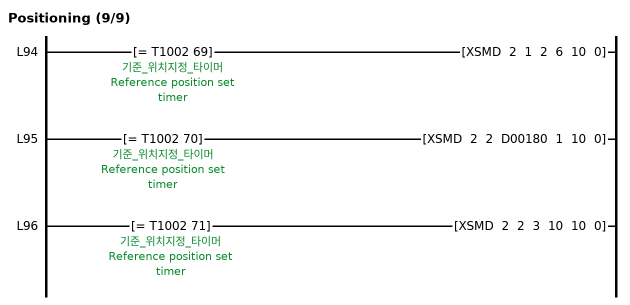
[picture p24: Positioning rungs L94-L96]
; L94
LOAD=     T1002 69	// 기준_위치지정_타이머 Reference position set timer
XSMD      2 1 2 6 10 0
; L95
LOAD=     T1002 70	// 기준_위치지정_타이머 Reference position set timer
XSMD      2 2 D00180 1 10 0
; L96
LOAD=     T1002 71	// 기준_위치지정_타이머 Reference position set timer
XSMD      2 2 3 10 10 0

PROGRAM PosItion_Switch (task: 스캔 프로그램)

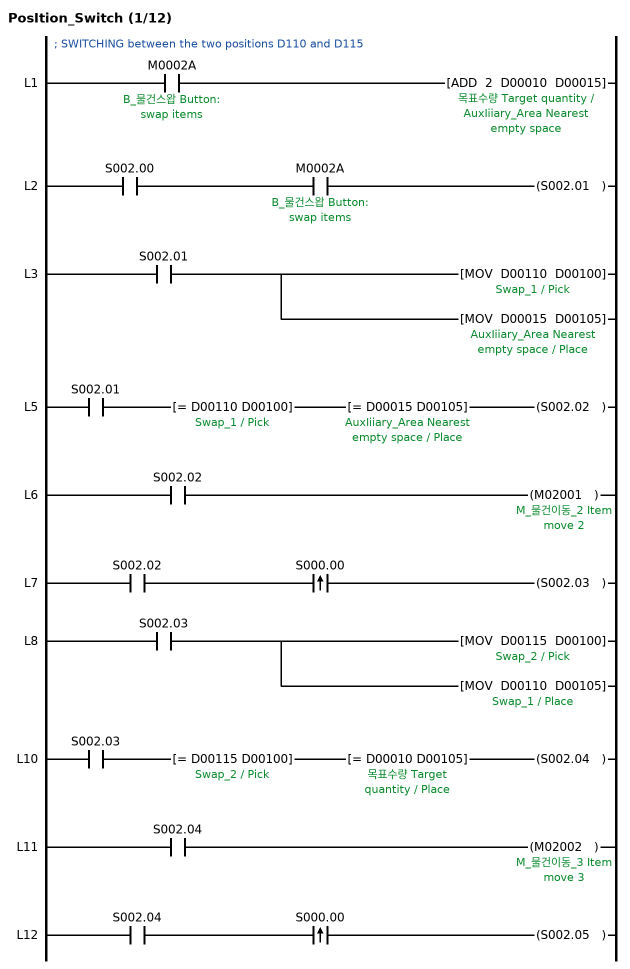
// SWITCHING between the two positions D110 and D115
; L1
LOAD      M0002A	// B_물건스왑 Button: swap items
ADD       2 D00010 D00015	// 목표수량 Target quantity / AuxIiiary_Area Nearest empty space
; L2
LOAD      S002.00
AND       M0002A	// B_물건스왑 Button: swap items
OUT       S002.01
; L3
LOAD      S002.01
MOV       D00110 D00100	// Swap_1 / Pick
MOV       D00015 D00105	// AuxIiiary_Area Nearest empty space / Place
; L5
LOAD      S002.01
AND=      D00110 D00100	// Swap_1 / Pick
AND=      D00015 D00105	// AuxIiiary_Area Nearest empty space / Place
OUT       S002.02
; L6
LOAD      S002.02
OUT       M02001	// M_물건이동_2 Item move 2
; L7
LOAD      S002.02
ANDP      S000.00
OUT       S002.03
; L8
LOAD      S002.03
MOV       D00115 D00100	// Swap_2 / Pick
MOV       D00110 D00105	// Swap_1 / Place
; L10
LOAD      S002.03
AND=      D00115 D00100	// Swap_2 / Pick
AND=      D00010 D00105	// 목표수량 Target quantity / Place
OUT       S002.04
; L11
LOAD      S002.04
OUT       M02002	// M_물건이동_3 Item move 3
; L12
LOAD      S002.04
ANDP      S000.00
OUT       S002.05

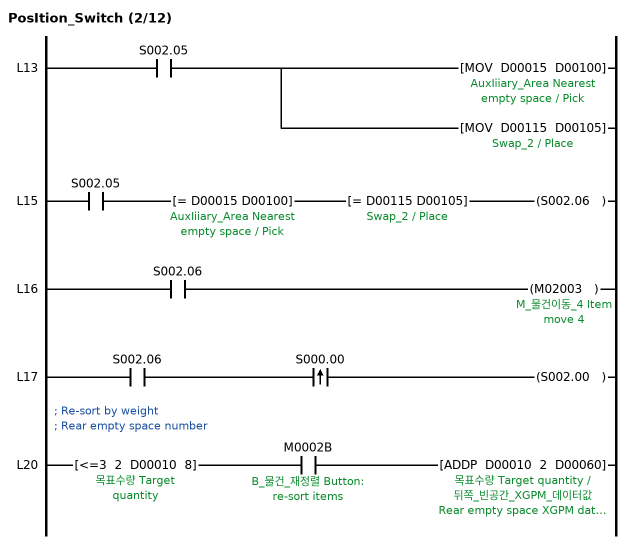
; L13
LOAD      S002.05
MOV       D00015 D00100	// AuxIiiary_Area Nearest empty space / Pick
MOV       D00115 D00105	// Swap_2 / Place
; L15
LOAD      S002.05
AND=      D00015 D00100	// AuxIiiary_Area Nearest empty space / Pick
AND=      D00115 D00105	// Swap_2 / Place
OUT       S002.06
; L16
LOAD      S002.06
OUT       M02003	// M_물건이동_4 Item move 4
; L17
LOAD      S002.06
ANDP      S000.00
OUT       S002.00
// Re-sort by weight
// Rear empty space number
; L20
LOAD<=3   2 D00010 8	// 목표수량 Target quantity
AND       M0002B	// B_물건_재정렬 Button: re-sort items
ADDP      D00010 2 D00060	// 목표수량 Target quantity / 뒤쪽_빈공간_XGPM_데이터값 Rear empty space XGPM data value

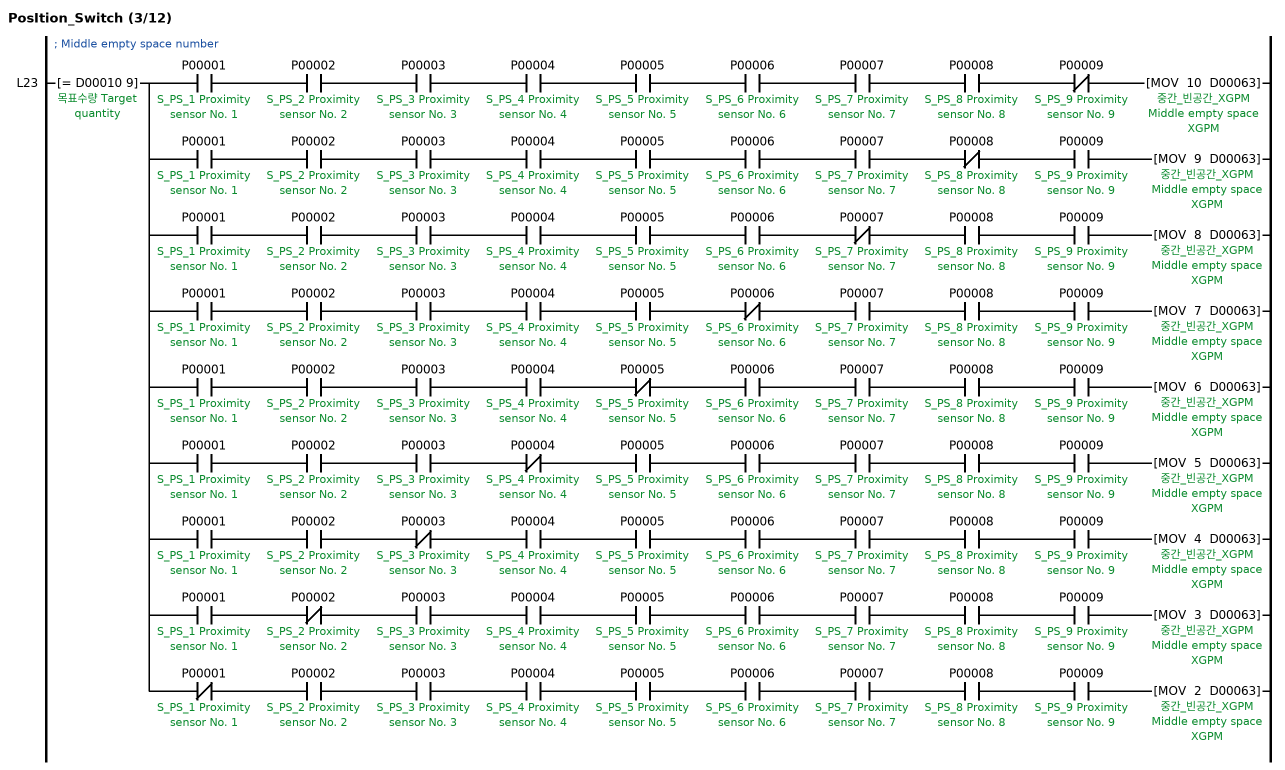
// Middle empty space number
; L23
LOAD=     D00010 9	// 목표수량 Target quantity
MPUSH
AND       P00001	// S_PS_1 Proximity sensor No. 1
AND       P00002	// S_PS_2 Proximity sensor No. 2
AND       P00003	// S_PS_3 Proximity sensor No. 3
AND       P00004	// S_PS_4 Proximity sensor No. 4
AND       P00005	// S_PS_5 Proximity sensor No. 5
AND       P00006	// S_PS_6 Proximity sensor No. 6
AND       P00007	// S_PS_7 Proximity sensor No. 7
AND       P00008	// S_PS_8 Proximity sensor No. 8
AND NOT   P00009	// S_PS_9 Proximity sensor No. 9
MOV       10 D00063	// 중간_빈공간_XGPM Middle empty space XGPM
MLOAD
AND       P00001	// S_PS_1 Proximity sensor No. 1
AND       P00002	// S_PS_2 Proximity sensor No. 2
AND       P00003	// S_PS_3 Proximity sensor No. 3
AND       P00004	// S_PS_4 Proximity sensor No. 4
AND       P00005	// S_PS_5 Proximity sensor No. 5
AND       P00006	// S_PS_6 Proximity sensor No. 6
AND       P00007	// S_PS_7 Proximity sensor No. 7
AND NOT   P00008	// S_PS_8 Proximity sensor No. 8
AND       P00009	// S_PS_9 Proximity sensor No. 9
MOV       9 D00063	// 중간_빈공간_XGPM Middle empty space XGPM
MLOAD
AND       P00001	// S_PS_1 Proximity sensor No. 1
AND       P00002	// S_PS_2 Proximity sensor No. 2
AND       P00003	// S_PS_3 Proximity sensor No. 3
AND       P00004	// S_PS_4 Proximity sensor No. 4
AND       P00005	// S_PS_5 Proximity sensor No. 5
AND       P00006	// S_PS_6 Proximity sensor No. 6
AND NOT   P00007	// S_PS_7 Proximity sensor No. 7
AND       P00008	// S_PS_8 Proximity sensor No. 8
AND       P00009	// S_PS_9 Proximity sensor No. 9
MOV       8 D00063	// 중간_빈공간_XGPM Middle empty space XGPM
MLOAD
AND       P00001	// S_PS_1 Proximity sensor No. 1
AND       P00002	// S_PS_2 Proximity sensor No. 2
AND       P00003	// S_PS_3 Proximity sensor No. 3
AND       P00004	// S_PS_4 Proximity sensor No. 4
AND       P00005	// S_PS_5 Proximity sensor No. 5
AND NOT   P00006	// S_PS_6 Proximity sensor No. 6
AND       P00007	// S_PS_7 Proximity sensor No. 7
AND       P00008	// S_PS_8 Proximity sensor No. 8
AND       P00009	// S_PS_9 Proximity sensor No. 9
MOV       7 D00063	// 중간_빈공간_XGPM Middle empty space XGPM
MLOAD
AND       P00001	// S_PS_1 Proximity sensor No. 1
AND       P00002	// S_PS_2 Proximity sensor No. 2
AND       P00003	// S_PS_3 Proximity sensor No. 3
AND       P00004	// S_PS_4 Proximity sensor No. 4
AND NOT   P00005	// S_PS_5 Proximity sensor No. 5
AND       P00006	// S_PS_6 Proximity sensor No. 6
AND       P00007	// S_PS_7 Proximity sensor No. 7
AND       P00008	// S_PS_8 Proximity sensor No. 8
AND       P00009	// S_PS_9 Proximity sensor No. 9
MOV       6 D00063	// 중간_빈공간_XGPM Middle empty space XGPM
MLOAD
AND       P00001	// S_PS_1 Proximity sensor No. 1
AND       P00002	// S_PS_2 Proximity sensor No. 2
AND       P00003	// S_PS_3 Proximity sensor No. 3
AND NOT   P00004	// S_PS_4 Proximity sensor No. 4
AND       P00005	// S_PS_5 Proximity sensor No. 5
AND       P00006	// S_PS_6 Proximity sensor No. 6
AND       P00007	// S_PS_7 Proximity sensor No. 7
AND       P00008	// S_PS_8 Proximity sensor No. 8
AND       P00009	// S_PS_9 Proximity sensor No. 9
MOV       5 D00063	// 중간_빈공간_XGPM Middle empty space XGPM
MLOAD
AND       P00001	// S_PS_1 Proximity sensor No. 1
AND       P00002	// S_PS_2 Proximity sensor No. 2
AND NOT   P00003	// S_PS_3 Proximity sensor No. 3
AND       P00004	// S_PS_4 Proximity sensor No. 4
AND       P00005	// S_PS_5 Proximity sensor No. 5
AND       P00006	// S_PS_6 Proximity sensor No. 6
AND       P00007	// S_PS_7 Proximity sensor No. 7
AND       P00008	// S_PS_8 Proximity sensor No. 8
AND       P00009	// S_PS_9 Proximity sensor No. 9
MOV       4 D00063	// 중간_빈공간_XGPM Middle empty space XGPM
MLOAD
AND       P00001	// S_PS_1 Proximity sensor No. 1
AND NOT   P00002	// S_PS_2 Proximity sensor No. 2
AND       P00003	// S_PS_3 Proximity sensor No. 3
AND       P00004	// S_PS_4 Proximity sensor No. 4
AND       P00005	// S_PS_5 Proximity sensor No. 5
AND       P00006	// S_PS_6 Proximity sensor No. 6
AND       P00007	// S_PS_7 Proximity sensor No. 7
AND       P00008	// S_PS_8 Proximity sensor No. 8
AND       P00009	// S_PS_9 Proximity sensor No. 9
MOV       3 D00063	// 중간_빈공간_XGPM Middle empty space XGPM
MPOP
AND NOT   P00001	// S_PS_1 Proximity sensor No. 1
AND       P00002	// S_PS_2 Proximity sensor No. 2
AND       P00003	// S_PS_3 Proximity sensor No. 3
AND       P00004	// S_PS_4 Proximity sensor No. 4
AND       P00005	// S_PS_5 Proximity sensor No. 5
AND       P00006	// S_PS_6 Proximity sensor No. 6
AND       P00007	// S_PS_7 Proximity sensor No. 7
AND       P00008	// S_PS_8 Proximity sensor No. 8
AND       P00009	// S_PS_9 Proximity sensor No. 9
MOV       2 D00063	// 중간_빈공간_XGPM Middle empty space XGPM

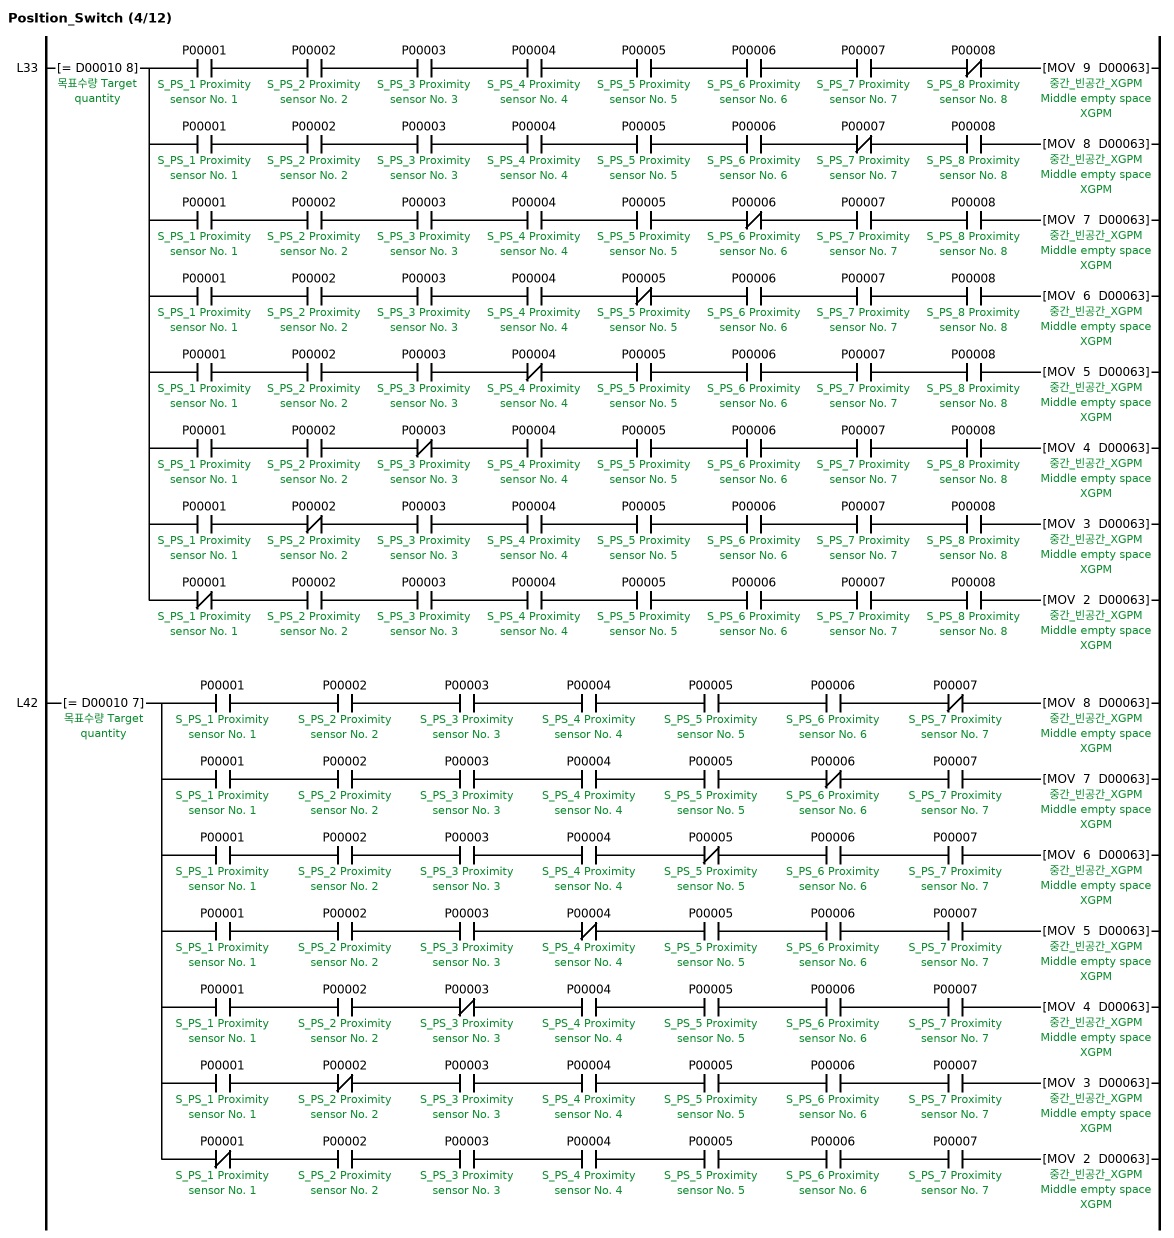
; L33
LOAD=     D00010 8	// 목표수량 Target quantity
MPUSH
AND       P00001	// S_PS_1 Proximity sensor No. 1
AND       P00002	// S_PS_2 Proximity sensor No. 2
AND       P00003	// S_PS_3 Proximity sensor No. 3
AND       P00004	// S_PS_4 Proximity sensor No. 4
AND       P00005	// S_PS_5 Proximity sensor No. 5
AND       P00006	// S_PS_6 Proximity sensor No. 6
AND       P00007	// S_PS_7 Proximity sensor No. 7
AND NOT   P00008	// S_PS_8 Proximity sensor No. 8
MOV       9 D00063	// 중간_빈공간_XGPM Middle empty space XGPM
MLOAD
AND       P00001	// S_PS_1 Proximity sensor No. 1
AND       P00002	// S_PS_2 Proximity sensor No. 2
AND       P00003	// S_PS_3 Proximity sensor No. 3
AND       P00004	// S_PS_4 Proximity sensor No. 4
AND       P00005	// S_PS_5 Proximity sensor No. 5
AND       P00006	// S_PS_6 Proximity sensor No. 6
AND NOT   P00007	// S_PS_7 Proximity sensor No. 7
AND       P00008	// S_PS_8 Proximity sensor No. 8
MOV       8 D00063	// 중간_빈공간_XGPM Middle empty space XGPM
MLOAD
AND       P00001	// S_PS_1 Proximity sensor No. 1
AND       P00002	// S_PS_2 Proximity sensor No. 2
AND       P00003	// S_PS_3 Proximity sensor No. 3
AND       P00004	// S_PS_4 Proximity sensor No. 4
AND       P00005	// S_PS_5 Proximity sensor No. 5
AND NOT   P00006	// S_PS_6 Proximity sensor No. 6
AND       P00007	// S_PS_7 Proximity sensor No. 7
AND       P00008	// S_PS_8 Proximity sensor No. 8
MOV       7 D00063	// 중간_빈공간_XGPM Middle empty space XGPM
MLOAD
AND       P00001	// S_PS_1 Proximity sensor No. 1
AND       P00002	// S_PS_2 Proximity sensor No. 2
AND       P00003	// S_PS_3 Proximity sensor No. 3
AND       P00004	// S_PS_4 Proximity sensor No. 4
AND NOT   P00005	// S_PS_5 Proximity sensor No. 5
AND       P00006	// S_PS_6 Proximity sensor No. 6
AND       P00007	// S_PS_7 Proximity sensor No. 7
AND       P00008	// S_PS_8 Proximity sensor No. 8
MOV       6 D00063	// 중간_빈공간_XGPM Middle empty space XGPM
MLOAD
AND       P00001	// S_PS_1 Proximity sensor No. 1
AND       P00002	// S_PS_2 Proximity sensor No. 2
AND       P00003	// S_PS_3 Proximity sensor No. 3
AND NOT   P00004	// S_PS_4 Proximity sensor No. 4
AND       P00005	// S_PS_5 Proximity sensor No. 5
AND       P00006	// S_PS_6 Proximity sensor No. 6
AND       P00007	// S_PS_7 Proximity sensor No. 7
AND       P00008	// S_PS_8 Proximity sensor No. 8
MOV       5 D00063	// 중간_빈공간_XGPM Middle empty space XGPM
MLOAD
AND       P00001	// S_PS_1 Proximity sensor No. 1
AND       P00002	// S_PS_2 Proximity sensor No. 2
AND NOT   P00003	// S_PS_3 Proximity sensor No. 3
AND       P00004	// S_PS_4 Proximity sensor No. 4
AND       P00005	// S_PS_5 Proximity sensor No. 5
AND       P00006	// S_PS_6 Proximity sensor No. 6
AND       P00007	// S_PS_7 Proximity sensor No. 7
AND       P00008	// S_PS_8 Proximity sensor No. 8
MOV       4 D00063	// 중간_빈공간_XGPM Middle empty space XGPM
MLOAD
AND       P00001	// S_PS_1 Proximity sensor No. 1
AND NOT   P00002	// S_PS_2 Proximity sensor No. 2
AND       P00003	// S_PS_3 Proximity sensor No. 3
AND       P00004	// S_PS_4 Proximity sensor No. 4
AND       P00005	// S_PS_5 Proximity sensor No. 5
AND       P00006	// S_PS_6 Proximity sensor No. 6
AND       P00007	// S_PS_7 Proximity sensor No. 7
AND       P00008	// S_PS_8 Proximity sensor No. 8
MOV       3 D00063	// 중간_빈공간_XGPM Middle empty space XGPM
MPOP
AND NOT   P00001	// S_PS_1 Proximity sensor No. 1
AND       P00002	// S_PS_2 Proximity sensor No. 2
AND       P00003	// S_PS_3 Proximity sensor No. 3
AND       P00004	// S_PS_4 Proximity sensor No. 4
AND       P00005	// S_PS_5 Proximity sensor No. 5
AND       P00006	// S_PS_6 Proximity sensor No. 6
AND       P00007	// S_PS_7 Proximity sensor No. 7
AND       P00008	// S_PS_8 Proximity sensor No. 8
MOV       2 D00063	// 중간_빈공간_XGPM Middle empty space XGPM
; L42
LOAD=     D00010 7	// 목표수량 Target quantity
MPUSH
AND       P00001	// S_PS_1 Proximity sensor No. 1
AND       P00002	// S_PS_2 Proximity sensor No. 2
AND       P00003	// S_PS_3 Proximity sensor No. 3
AND       P00004	// S_PS_4 Proximity sensor No. 4
AND       P00005	// S_PS_5 Proximity sensor No. 5
AND       P00006	// S_PS_6 Proximity sensor No. 6
AND NOT   P00007	// S_PS_7 Proximity sensor No. 7
MOV       8 D00063	// 중간_빈공간_XGPM Middle empty space XGPM
MLOAD
AND       P00001	// S_PS_1 Proximity sensor No. 1
AND       P00002	// S_PS_2 Proximity sensor No. 2
AND       P00003	// S_PS_3 Proximity sensor No. 3
AND       P00004	// S_PS_4 Proximity sensor No. 4
AND       P00005	// S_PS_5 Proximity sensor No. 5
AND NOT   P00006	// S_PS_6 Proximity sensor No. 6
AND       P00007	// S_PS_7 Proximity sensor No. 7
MOV       7 D00063	// 중간_빈공간_XGPM Middle empty space XGPM
MLOAD
AND       P00001	// S_PS_1 Proximity sensor No. 1
AND       P00002	// S_PS_2 Proximity sensor No. 2
AND       P00003	// S_PS_3 Proximity sensor No. 3
AND       P00004	// S_PS_4 Proximity sensor No. 4
AND NOT   P00005	// S_PS_5 Proximity sensor No. 5
AND       P00006	// S_PS_6 Proximity sensor No. 6
AND       P00007	// S_PS_7 Proximity sensor No. 7
MOV       6 D00063	// 중간_빈공간_XGPM Middle empty space XGPM
MLOAD
AND       P00001	// S_PS_1 Proximity sensor No. 1
AND       P00002	// S_PS_2 Proximity sensor No. 2
AND       P00003	// S_PS_3 Proximity sensor No. 3
AND NOT   P00004	// S_PS_4 Proximity sensor No. 4
AND       P00005	// S_PS_5 Proximity sensor No. 5
AND       P00006	// S_PS_6 Proximity sensor No. 6
AND       P00007	// S_PS_7 Proximity sensor No. 7
MOV       5 D00063	// 중간_빈공간_XGPM Middle empty space XGPM
MLOAD
AND       P00001	// S_PS_1 Proximity sensor No. 1
AND       P00002	// S_PS_2 Proximity sensor No. 2
AND NOT   P00003	// S_PS_3 Proximity sensor No. 3
AND       P00004	// S_PS_4 Proximity sensor No. 4
AND       P00005	// S_PS_5 Proximity sensor No. 5
AND       P00006	// S_PS_6 Proximity sensor No. 6
AND       P00007	// S_PS_7 Proximity sensor No. 7
MOV       4 D00063	// 중간_빈공간_XGPM Middle empty space XGPM
MLOAD
AND       P00001	// S_PS_1 Proximity sensor No. 1
AND NOT   P00002	// S_PS_2 Proximity sensor No. 2
AND       P00003	// S_PS_3 Proximity sensor No. 3
AND       P00004	// S_PS_4 Proximity sensor No. 4
AND       P00005	// S_PS_5 Proximity sensor No. 5
AND       P00006	// S_PS_6 Proximity sensor No. 6
AND       P00007	// S_PS_7 Proximity sensor No. 7
MOV       3 D00063	// 중간_빈공간_XGPM Middle empty space XGPM
MPOP
AND NOT   P00001	// S_PS_1 Proximity sensor No. 1
AND       P00002	// S_PS_2 Proximity sensor No. 2
AND       P00003	// S_PS_3 Proximity sensor No. 3
AND       P00004	// S_PS_4 Proximity sensor No. 4
AND       P00005	// S_PS_5 Proximity sensor No. 5
AND       P00006	// S_PS_6 Proximity sensor No. 6
AND       P00007	// S_PS_7 Proximity sensor No. 7
MOV       2 D00063	// 중간_빈공간_XGPM Middle empty space XGPM

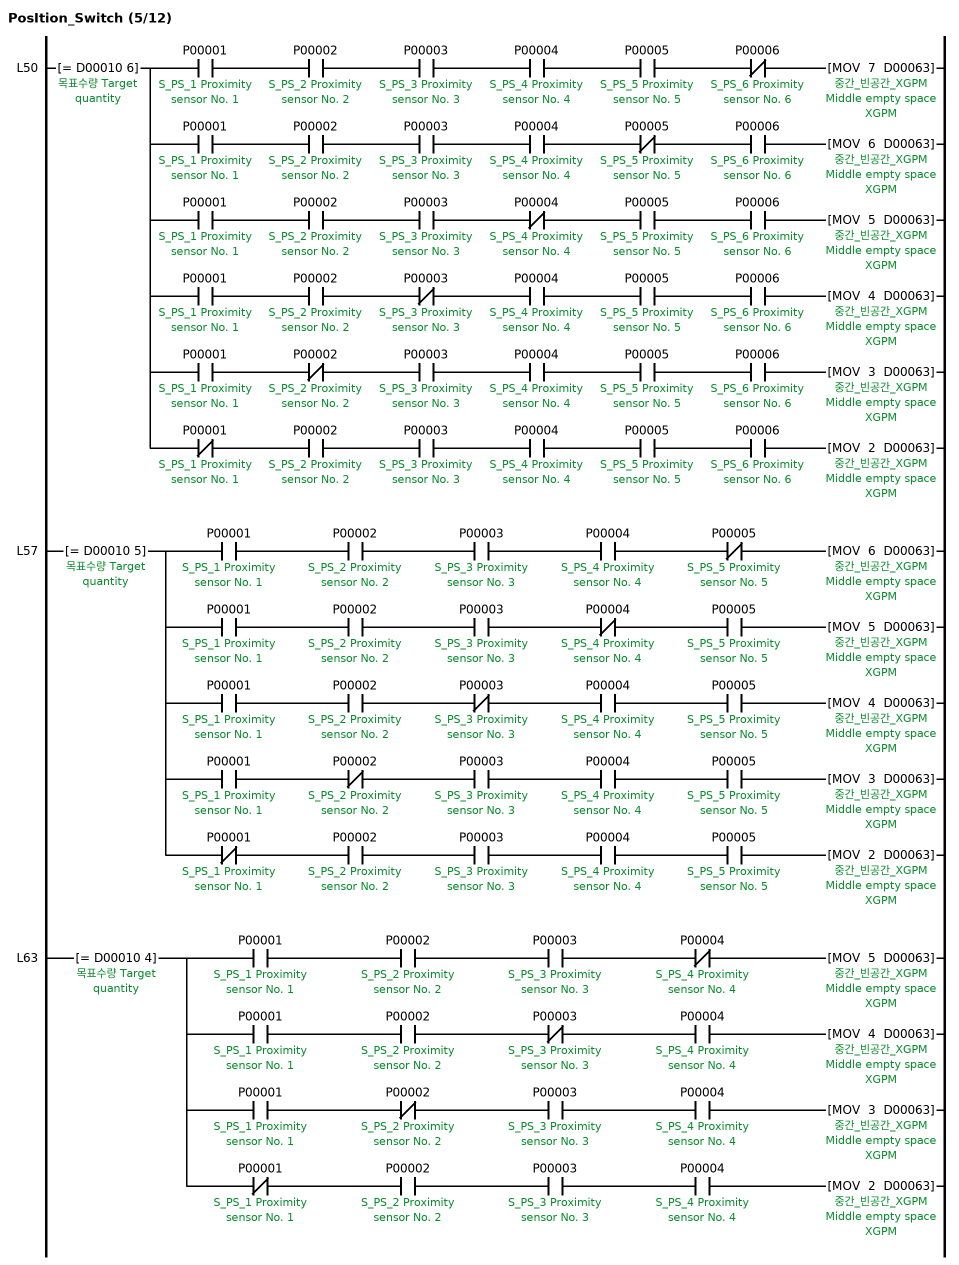
; L50
LOAD=     D00010 6	// 목표수량 Target quantity
MPUSH
AND       P00001	// S_PS_1 Proximity sensor No. 1
AND       P00002	// S_PS_2 Proximity sensor No. 2
AND       P00003	// S_PS_3 Proximity sensor No. 3
AND       P00004	// S_PS_4 Proximity sensor No. 4
AND       P00005	// S_PS_5 Proximity sensor No. 5
AND NOT   P00006	// S_PS_6 Proximity sensor No. 6
MOV       7 D00063	// 중간_빈공간_XGPM Middle empty space XGPM
MLOAD
AND       P00001	// S_PS_1 Proximity sensor No. 1
AND       P00002	// S_PS_2 Proximity sensor No. 2
AND       P00003	// S_PS_3 Proximity sensor No. 3
AND       P00004	// S_PS_4 Proximity sensor No. 4
AND NOT   P00005	// S_PS_5 Proximity sensor No. 5
AND       P00006	// S_PS_6 Proximity sensor No. 6
MOV       6 D00063	// 중간_빈공간_XGPM Middle empty space XGPM
MLOAD
AND       P00001	// S_PS_1 Proximity sensor No. 1
AND       P00002	// S_PS_2 Proximity sensor No. 2
AND       P00003	// S_PS_3 Proximity sensor No. 3
AND NOT   P00004	// S_PS_4 Proximity sensor No. 4
AND       P00005	// S_PS_5 Proximity sensor No. 5
AND       P00006	// S_PS_6 Proximity sensor No. 6
MOV       5 D00063	// 중간_빈공간_XGPM Middle empty space XGPM
MLOAD
AND       P00001	// S_PS_1 Proximity sensor No. 1
AND       P00002	// S_PS_2 Proximity sensor No. 2
AND NOT   P00003	// S_PS_3 Proximity sensor No. 3
AND       P00004	// S_PS_4 Proximity sensor No. 4
AND       P00005	// S_PS_5 Proximity sensor No. 5
AND       P00006	// S_PS_6 Proximity sensor No. 6
MOV       4 D00063	// 중간_빈공간_XGPM Middle empty space XGPM
MLOAD
AND       P00001	// S_PS_1 Proximity sensor No. 1
AND NOT   P00002	// S_PS_2 Proximity sensor No. 2
AND       P00003	// S_PS_3 Proximity sensor No. 3
AND       P00004	// S_PS_4 Proximity sensor No. 4
AND       P00005	// S_PS_5 Proximity sensor No. 5
AND       P00006	// S_PS_6 Proximity sensor No. 6
MOV       3 D00063	// 중간_빈공간_XGPM Middle empty space XGPM
MPOP
AND NOT   P00001	// S_PS_1 Proximity sensor No. 1
AND       P00002	// S_PS_2 Proximity sensor No. 2
AND       P00003	// S_PS_3 Proximity sensor No. 3
AND       P00004	// S_PS_4 Proximity sensor No. 4
AND       P00005	// S_PS_5 Proximity sensor No. 5
AND       P00006	// S_PS_6 Proximity sensor No. 6
MOV       2 D00063	// 중간_빈공간_XGPM Middle empty space XGPM
; L57
LOAD=     D00010 5	// 목표수량 Target quantity
MPUSH
AND       P00001	// S_PS_1 Proximity sensor No. 1
AND       P00002	// S_PS_2 Proximity sensor No. 2
AND       P00003	// S_PS_3 Proximity sensor No. 3
AND       P00004	// S_PS_4 Proximity sensor No. 4
AND NOT   P00005	// S_PS_5 Proximity sensor No. 5
MOV       6 D00063	// 중간_빈공간_XGPM Middle empty space XGPM
MLOAD
AND       P00001	// S_PS_1 Proximity sensor No. 1
AND       P00002	// S_PS_2 Proximity sensor No. 2
AND       P00003	// S_PS_3 Proximity sensor No. 3
AND NOT   P00004	// S_PS_4 Proximity sensor No. 4
AND       P00005	// S_PS_5 Proximity sensor No. 5
MOV       5 D00063	// 중간_빈공간_XGPM Middle empty space XGPM
MLOAD
AND       P00001	// S_PS_1 Proximity sensor No. 1
AND       P00002	// S_PS_2 Proximity sensor No. 2
AND NOT   P00003	// S_PS_3 Proximity sensor No. 3
AND       P00004	// S_PS_4 Proximity sensor No. 4
AND       P00005	// S_PS_5 Proximity sensor No. 5
MOV       4 D00063	// 중간_빈공간_XGPM Middle empty space XGPM
MLOAD
AND       P00001	// S_PS_1 Proximity sensor No. 1
AND NOT   P00002	// S_PS_2 Proximity sensor No. 2
AND       P00003	// S_PS_3 Proximity sensor No. 3
AND       P00004	// S_PS_4 Proximity sensor No. 4
AND       P00005	// S_PS_5 Proximity sensor No. 5
MOV       3 D00063	// 중간_빈공간_XGPM Middle empty space XGPM
MPOP
AND NOT   P00001	// S_PS_1 Proximity sensor No. 1
AND       P00002	// S_PS_2 Proximity sensor No. 2
AND       P00003	// S_PS_3 Proximity sensor No. 3
AND       P00004	// S_PS_4 Proximity sensor No. 4
AND       P00005	// S_PS_5 Proximity sensor No. 5
MOV       2 D00063	// 중간_빈공간_XGPM Middle empty space XGPM
; L63
LOAD=     D00010 4	// 목표수량 Target quantity
MPUSH
AND       P00001	// S_PS_1 Proximity sensor No. 1
AND       P00002	// S_PS_2 Proximity sensor No. 2
AND       P00003	// S_PS_3 Proximity sensor No. 3
AND NOT   P00004	// S_PS_4 Proximity sensor No. 4
MOV       5 D00063	// 중간_빈공간_XGPM Middle empty space XGPM
MLOAD
AND       P00001	// S_PS_1 Proximity sensor No. 1
AND       P00002	// S_PS_2 Proximity sensor No. 2
AND NOT   P00003	// S_PS_3 Proximity sensor No. 3
AND       P00004	// S_PS_4 Proximity sensor No. 4
MOV       4 D00063	// 중간_빈공간_XGPM Middle empty space XGPM
MLOAD
AND       P00001	// S_PS_1 Proximity sensor No. 1
AND NOT   P00002	// S_PS_2 Proximity sensor No. 2
AND       P00003	// S_PS_3 Proximity sensor No. 3
AND       P00004	// S_PS_4 Proximity sensor No. 4
MOV       3 D00063	// 중간_빈공간_XGPM Middle empty space XGPM
MPOP
AND NOT   P00001	// S_PS_1 Proximity sensor No. 1
AND       P00002	// S_PS_2 Proximity sensor No. 2
AND       P00003	// S_PS_3 Proximity sensor No. 3
AND       P00004	// S_PS_4 Proximity sensor No. 4
MOV       2 D00063	// 중간_빈공간_XGPM Middle empty space XGPM

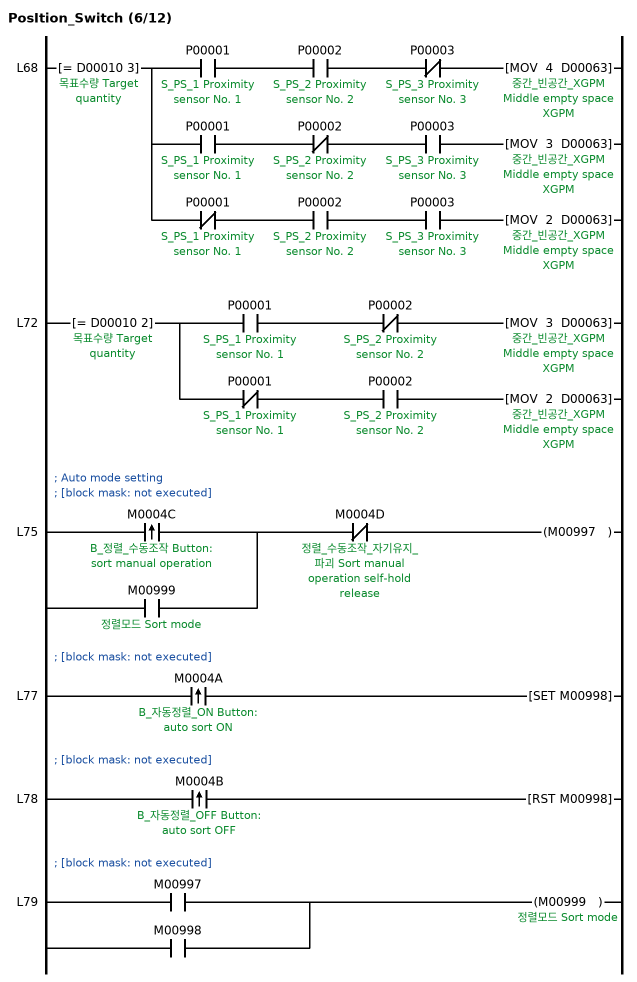
; L68
LOAD=     D00010 3	// 목표수량 Target quantity
MPUSH
AND       P00001	// S_PS_1 Proximity sensor No. 1
AND       P00002	// S_PS_2 Proximity sensor No. 2
AND NOT   P00003	// S_PS_3 Proximity sensor No. 3
MOV       4 D00063	// 중간_빈공간_XGPM Middle empty space XGPM
MLOAD
AND       P00001	// S_PS_1 Proximity sensor No. 1
AND NOT   P00002	// S_PS_2 Proximity sensor No. 2
AND       P00003	// S_PS_3 Proximity sensor No. 3
MOV       3 D00063	// 중간_빈공간_XGPM Middle empty space XGPM
MPOP
AND NOT   P00001	// S_PS_1 Proximity sensor No. 1
AND       P00002	// S_PS_2 Proximity sensor No. 2
AND       P00003	// S_PS_3 Proximity sensor No. 3
MOV       2 D00063	// 중간_빈공간_XGPM Middle empty space XGPM
; L72
LOAD=     D00010 2	// 목표수량 Target quantity
MPUSH
AND       P00001	// S_PS_1 Proximity sensor No. 1
AND NOT   P00002	// S_PS_2 Proximity sensor No. 2
MOV       3 D00063	// 중간_빈공간_XGPM Middle empty space XGPM
MPOP
AND NOT   P00001	// S_PS_1 Proximity sensor No. 1
AND       P00002	// S_PS_2 Proximity sensor No. 2
MOV       2 D00063	// 중간_빈공간_XGPM Middle empty space XGPM
// Auto mode setting
; L75 (block mask: not executed)
LOADP     M0004C	// B_정렬_수동조작 Button: sort manual operation
OR        M00999	// 정렬모드 Sort mode
AND NOT   M0004D	// 정렬_수동조작_자기유지_파괴 Sort manual operation self-hold release
OUT       M00997
; L77 (block mask: not executed)
LOADP     M0004A	// B_자동정렬_ON Button: auto sort ON
SET       M00998
; L78 (block mask: not executed)
LOADP     M0004B	// B_자동정렬_OFF Button: auto sort OFF
RST       M00998
; L79 (block mask: not executed)
LOAD      M00997
OR        M00998
OUT       M00999	// 정렬모드 Sort mode

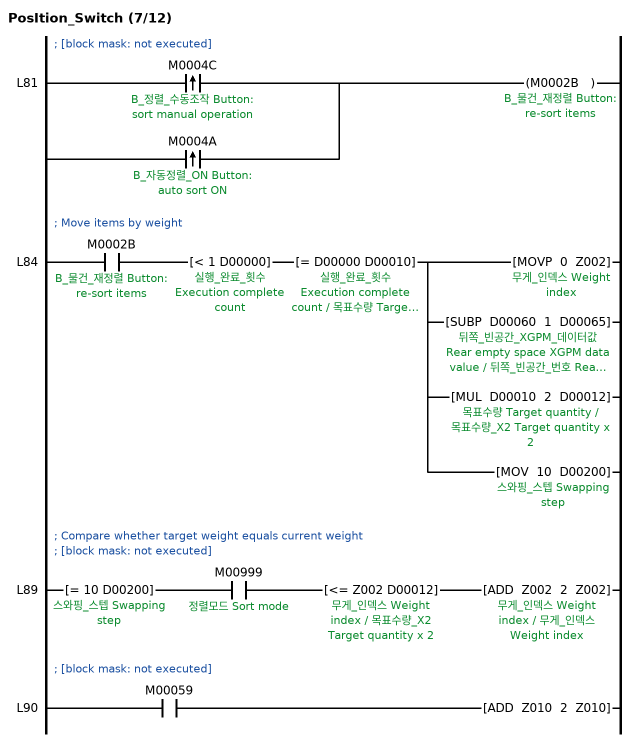
; L81 (block mask: not executed)
LOADP     M0004C	// B_정렬_수동조작 Button: sort manual operation
ORP       M0004A	// B_자동정렬_ON Button: auto sort ON
OUT       M0002B	// B_물건_재정렬 Button: re-sort items
// Move items by weight
; L84
LOAD      M0002B	// B_물건_재정렬 Button: re-sort items
AND<      1 D00000	// 실행_완료_횟수 Execution complete count
AND=      D00000 D00010	// 실행_완료_횟수 Execution complete count / 목표수량 Target quantity
MOVP      0 Z002	// 무게_인덱스 Weight index
SUBP      D00060 1 D00065	// 뒤쪽_빈공간_XGPM_데이터값 Rear empty space XGPM data value / 뒤쪽_빈공간_번호 Rear empty space number
MUL       D00010 2 D00012	// 목표수량 Target quantity / 목표수량_X2 Target quantity x 2
MOV       10 D00200	// 스와핑_스텝 Swapping step
// Compare whether target weight equals current weight
; L89 (block mask: not executed)
LOAD=     10 D00200	// 스와핑_스텝 Swapping step
AND       M00999	// 정렬모드 Sort mode
AND<=     Z002 D00012	// 무게_인덱스 Weight index / 목표수량_X2 Target quantity x 2
ADD       Z002 2 Z002	// 무게_인덱스 Weight index / 무게_인덱스 Weight index
; L90 (block mask: not executed)
LOAD      M00059
ADD       Z010 2 Z010

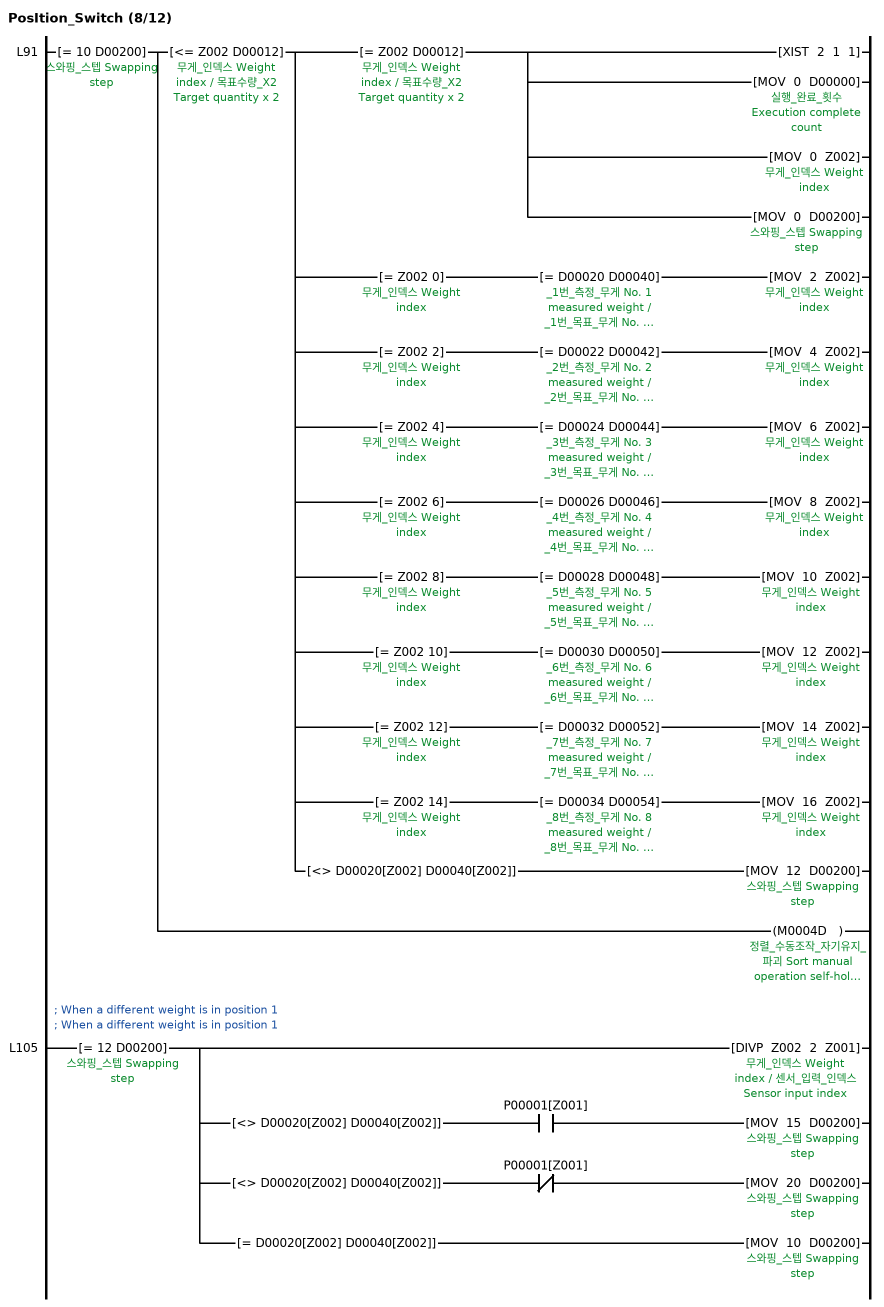
; L91
LOAD=     10 D00200	// 스와핑_스텝 Swapping step
MPUSH
AND<=     Z002 D00012	// 무게_인덱스 Weight index / 목표수량_X2 Target quantity x 2
MPUSH
AND=      Z002 D00012	// 무게_인덱스 Weight index / 목표수량_X2 Target quantity x 2
XIST      2 1 1
MOV       0 D00000	// 실행_완료_횟수 Execution complete count
MOV       0 Z002	// 무게_인덱스 Weight index
MOV       0 D00200	// 스와핑_스텝 Swapping step
MLOAD
AND=      Z002 0	// 무게_인덱스 Weight index
AND=      D00020 D00040	// _1번_측정_무게 No. 1 measured weight / _1번_목표_무게 No. 1 target weight
MOV       2 Z002	// 무게_인덱스 Weight index
MLOAD
AND=      Z002 2	// 무게_인덱스 Weight index
AND=      D00022 D00042	// _2번_측정_무게 No. 2 measured weight / _2번_목표_무게 No. 2 target weight
MOV       4 Z002	// 무게_인덱스 Weight index
MLOAD
AND=      Z002 4	// 무게_인덱스 Weight index
AND=      D00024 D00044	// _3번_측정_무게 No. 3 measured weight / _3번_목표_무게 No. 3 target weight
MOV       6 Z002	// 무게_인덱스 Weight index
MLOAD
AND=      Z002 6	// 무게_인덱스 Weight index
AND=      D00026 D00046	// _4번_측정_무게 No. 4 measured weight / _4번_목표_무게 No. 4 target weight
MOV       8 Z002	// 무게_인덱스 Weight index
MLOAD
AND=      Z002 8	// 무게_인덱스 Weight index
AND=      D00028 D00048	// _5번_측정_무게 No. 5 measured weight / _5번_목표_무게 No. 5 target weight
MOV       10 Z002	// 무게_인덱스 Weight index
MLOAD
AND=      Z002 10	// 무게_인덱스 Weight index
AND=      D00030 D00050	// _6번_측정_무게 No. 6 measured weight / _6번_목표_무게 No. 6 target weight
MOV       12 Z002	// 무게_인덱스 Weight index
MLOAD
AND=      Z002 12	// 무게_인덱스 Weight index
AND=      D00032 D00052	// _7번_측정_무게 No. 7 measured weight / _7번_목표_무게 No. 7 target weight
MOV       14 Z002	// 무게_인덱스 Weight index
MLOAD
AND=      Z002 14	// 무게_인덱스 Weight index
AND=      D00034 D00054	// _8번_측정_무게 No. 8 measured weight / _8번_목표_무게 No. 8 target weight
MOV       16 Z002	// 무게_인덱스 Weight index
MPOP
AND<>     D00020[Z002] D00040[Z002]
MOV       12 D00200	// 스와핑_스텝 Swapping step
MPOP
OUT       M0004D	// 정렬_수동조작_자기유지_파괴 Sort manual operation self-hold release
; L105
LOAD=     12 D00200	// 스와핑_스텝 Swapping step
DIVP      Z002 2 Z001	// 무게_인덱스 Weight index / 센서_입력_인덱스 Sensor input index
MPUSH
AND<>     D00020[Z002] D00040[Z002]
AND       P00001[Z001]
MOV       15 D00200	// 스와핑_스텝 Swapping step
MLOAD
AND<>     D00020[Z002] D00040[Z002]
AND NOT   P00001[Z001]
MOV       20 D00200	// 스와핑_스텝 Swapping step
MPOP
AND=      D00020[Z002] D00040[Z002]
MOV       10 D00200	// 스와핑_스텝 Swapping step
// output comment: When a different weight is in position 1
// output comment: When a different weight is in position 1

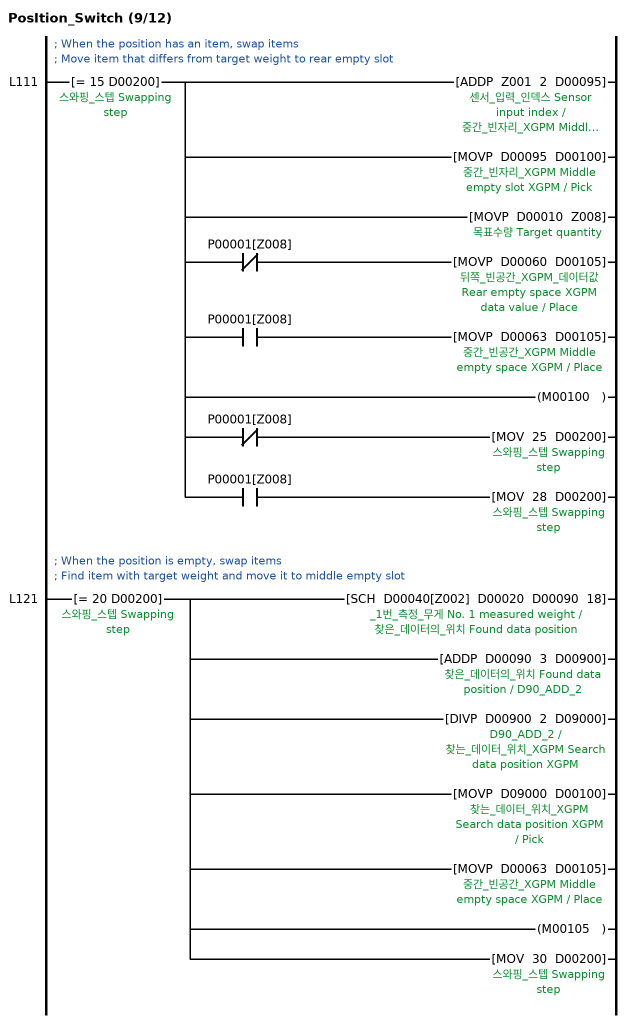
// When the position has an item, swap items
// Move item that differs from target weight to rear empty slot
; L111
LOAD=     15 D00200	// 스와핑_스텝 Swapping step
ADDP      Z001 2 D00095	// 센서_입력_인덱스 Sensor input index / 중간_빈자리_XGPM Middle empty slot XGPM
MOVP      D00095 D00100	// 중간_빈자리_XGPM Middle empty slot XGPM / Pick
MOVP      D00010 Z008	// 목표수량 Target quantity
MPUSH
AND NOT   P00001[Z008]
MOVP      D00060 D00105	// 뒤쪽_빈공간_XGPM_데이터값 Rear empty space XGPM data value / Place
MLOAD
AND       P00001[Z008]
MOVP      D00063 D00105	// 중간_빈공간_XGPM Middle empty space XGPM / Place
MLOAD
OUT       M00100
AND NOT   P00001[Z008]
MOV       25 D00200	// 스와핑_스텝 Swapping step
MPOP
AND       P00001[Z008]
MOV       28 D00200	// 스와핑_스텝 Swapping step
// When the position is empty, swap items
// Find item with target weight and move it to middle empty slot
; L121
LOAD=     20 D00200	// 스와핑_스텝 Swapping step
SCH       D00040[Z002] D00020 D00090 18	// _1번_측정_무게 No. 1 measured weight / 찾은_데이터의_위치 Found data position
ADDP      D00090 3 D00900	// 찾은_데이터의_위치 Found data position / D90_ADD_2
DIVP      D00900 2 D09000	// D90_ADD_2 / 찾는_데이터_위치_XGPM Search data position XGPM
MOVP      D09000 D00100	// 찾는_데이터_위치_XGPM Search data position XGPM / Pick
MOVP      D00063 D00105	// 중간_빈공간_XGPM Middle empty space XGPM / Place
OUT       M00105
MOV       30 D00200	// 스와핑_스텝 Swapping step

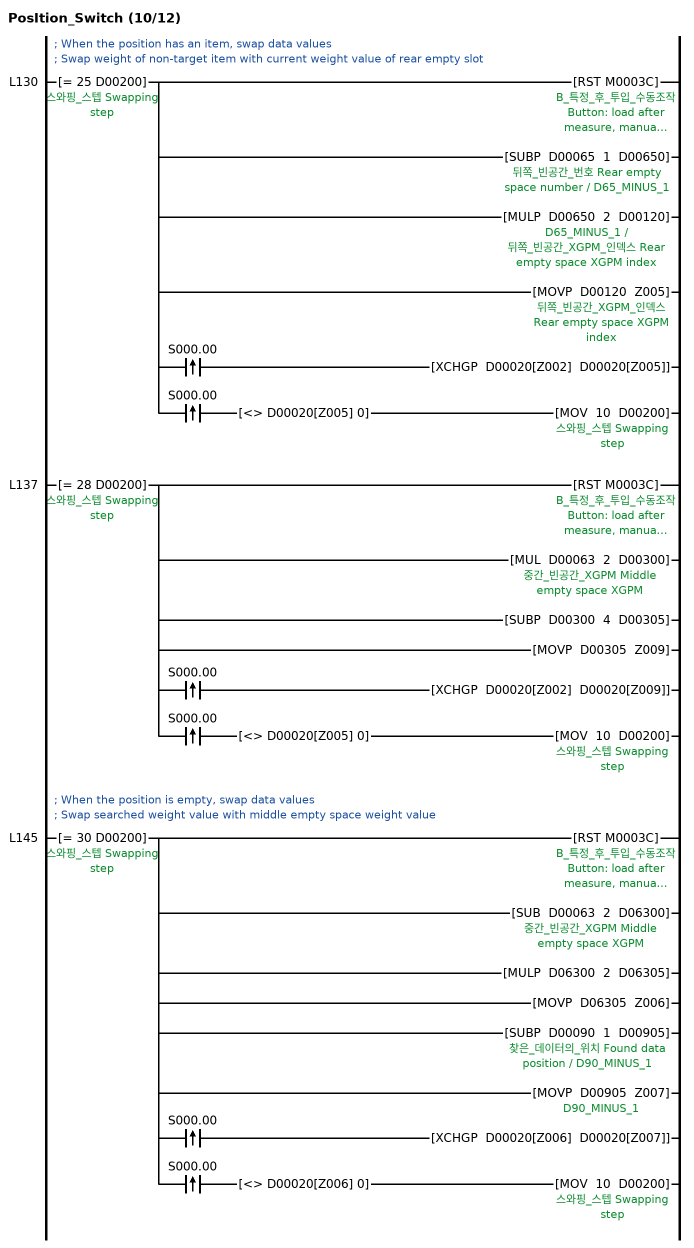
// When the position has an item, swap data values
// Swap weight of non-target item with current weight value of rear empty slot
; L130
LOAD=     25 D00200	// 스와핑_스텝 Swapping step
RST       M0003C	// B_특정_후_투입_수동조작 Button: load after measure, manual operation
SUBP      D00065 1 D00650	// 뒤쪽_빈공간_번호 Rear empty space number / D65_MINUS_1
MULP      D00650 2 D00120	// D65_MINUS_1 / 뒤쪽_빈공간_XGPM_인덱스 Rear empty space XGPM index
MOVP      D00120 Z005	// 뒤쪽_빈공간_XGPM_인덱스 Rear empty space XGPM index
MPUSH
ANDP      S000.00
XCHGP     D00020[Z002] D00020[Z005]
MPOP
ANDP      S000.00
AND<>     D00020[Z005] 0
MOV       10 D00200	// 스와핑_스텝 Swapping step
; L137
LOAD=     28 D00200	// 스와핑_스텝 Swapping step
RST       M0003C	// B_특정_후_투입_수동조작 Button: load after measure, manual operation
MUL       D00063 2 D00300	// 중간_빈공간_XGPM Middle empty space XGPM
SUBP      D00300 4 D00305
MOVP      D00305 Z009
MPUSH
ANDP      S000.00
XCHGP     D00020[Z002] D00020[Z009]
MPOP
ANDP      S000.00
AND<>     D00020[Z005] 0
MOV       10 D00200	// 스와핑_스텝 Swapping step
// When the position is empty, swap data values
// Swap searched weight value with middle empty space weight value
; L145
LOAD=     30 D00200	// 스와핑_스텝 Swapping step
RST       M0003C	// B_특정_후_투입_수동조작 Button: load after measure, manual operation
SUB       D00063 2 D06300	// 중간_빈공간_XGPM Middle empty space XGPM
MULP      D06300 2 D06305
MOVP      D06305 Z006
SUBP      D00090 1 D00905	// 찾은_데이터의_위치 Found data position / D90_MINUS_1
MOVP      D00905 Z007	// D90_MINUS_1
MPUSH
ANDP      S000.00
XCHGP     D00020[Z006] D00020[Z007]
MPOP
ANDP      S000.00
AND<>     D00020[Z006] 0
MOV       10 D00200	// 스와핑_스텝 Swapping step

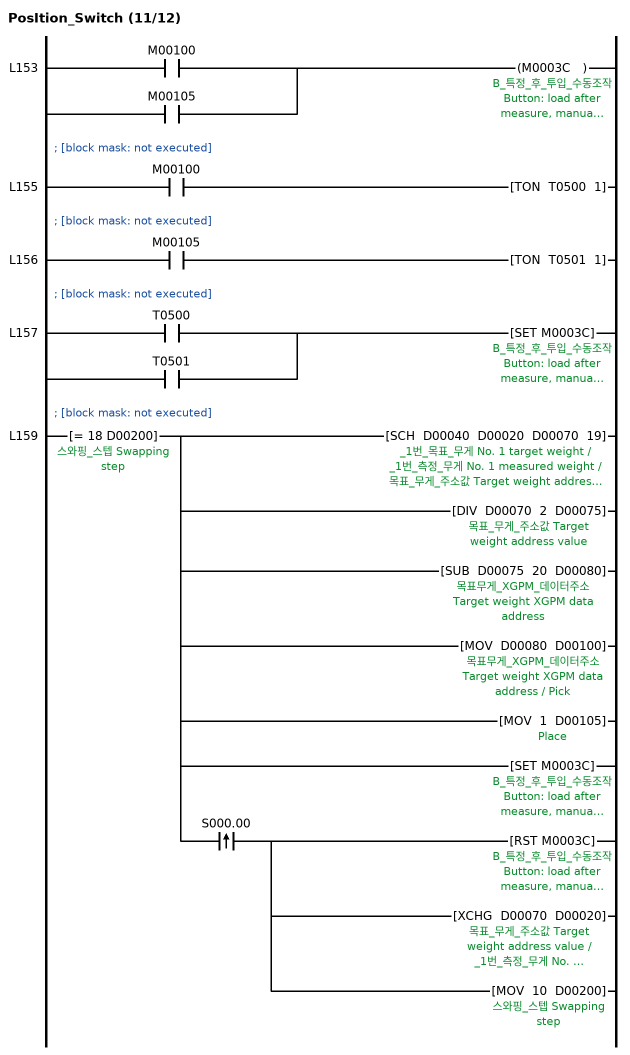
; L153
LOAD      M00100
OR        M00105
OUT       M0003C	// B_특정_후_투입_수동조작 Button: load after measure, manual operation
; L155 (block mask: not executed)
LOAD      M00100
TON       T0500 1
; L156 (block mask: not executed)
LOAD      M00105
TON       T0501 1
; L157 (block mask: not executed)
LOAD      T0500
OR        T0501
SET       M0003C	// B_특정_후_투입_수동조작 Button: load after measure, manual operation
; L159 (block mask: not executed)
LOAD=     18 D00200	// 스와핑_스텝 Swapping step
SCH       D00040 D00020 D00070 19	// _1번_목표_무게 No. 1 target weight / _1번_측정_무게 No. 1 measured weight / 목표_무게_주소값 Target weight address value
DIV       D00070 2 D00075	// 목표_무게_주소값 Target weight address value
SUB       D00075 20 D00080	// 목표무게_XGPM_데이터주소 Target weight XGPM data address
MOV       D00080 D00100	// 목표무게_XGPM_데이터주소 Target weight XGPM data address / Pick
MOV       1 D00105	// Place
SET       M0003C	// B_특정_후_투입_수동조작 Button: load after measure, manual operation
ANDP      S000.00
RST       M0003C	// B_특정_후_투입_수동조작 Button: load after measure, manual operation
XCHG      D00070 D00020	// 목표_무게_주소값 Target weight address value / _1번_측정_무게 No. 1 measured weight
MOV       10 D00200	// 스와핑_스텝 Swapping step

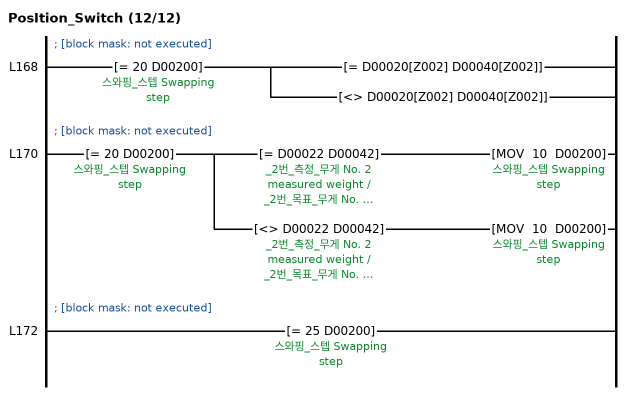
; L168 (block mask: not executed)
LOAD=     20 D00200	// 스와핑_스텝 Swapping step
LOAD=     D00020[Z002] D00040[Z002]
OR<>      D00020[Z002] D00040[Z002]
AND LOAD
; L170 (block mask: not executed)
LOAD=     20 D00200	// 스와핑_스텝 Swapping step
MPUSH
AND=      D00022 D00042	// _2번_측정_무게 No. 2 measured weight / _2번_목표_무게 No. 2 target weight
MOV       10 D00200	// 스와핑_스텝 Swapping step
MPOP
AND<>     D00022 D00042	// _2번_측정_무게 No. 2 measured weight / _2번_목표_무게 No. 2 target weight
MOV       10 D00200	// 스와핑_스텝 Swapping step
; L172 (block mask: not executed)
LOAD=     25 D00200	// 스와핑_스텝 Swapping step

PROGRAM Operation (task: 스캔 프로그램)

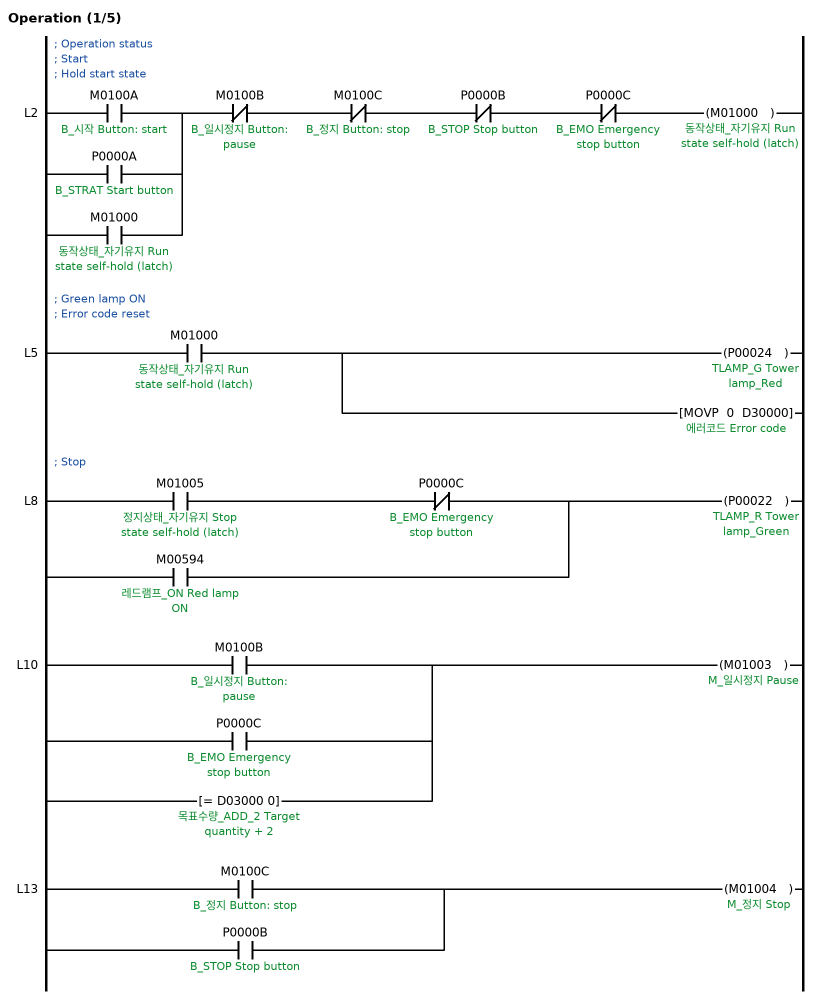
// Operation status
// Start
; L2
LOAD      M0100A	// B_시작 Button: start
OR        P0000A	// B_STRAT Start button
OR        M01000	// 동작상태_자기유지 Run state self-hold (latch)
AND NOT   M0100B	// B_일시정지 Button: pause
AND NOT   M0100C	// B_정지 Button: stop
AND NOT   P0000B	// B_STOP Stop button
AND NOT   P0000C	// B_EMO Emergency stop button
OUT       M01000	// 동작상태_자기유지 Run state self-hold (latch)
// output comment: Hold start state
; L5
LOAD      M01000	// 동작상태_자기유지 Run state self-hold (latch)
OUT       P00024	// TLAMP_G Tower lamp_Red
MOVP      0 D30000	// 에러코드 Error code
// output comment: Green lamp ON
// output comment: Error code reset
// Stop
; L8
LOAD      M01005	// 정지상태_자기유지 Stop state self-hold (latch)
AND NOT   P0000C	// B_EMO Emergency stop button
OR        M00594	// 레드램프_ON Red lamp ON
OUT       P00022	// TLAMP_R Tower lamp_Green
; L10
LOAD      M0100B	// B_일시정지 Button: pause
OR        P0000C	// B_EMO Emergency stop button
OR=       D03000 0	// 목표수량_ADD_2 Target quantity + 2
OUT       M01003	// M_일시정지 Pause
; L13
LOAD      M0100C	// B_정지 Button: stop
OR        P0000B	// B_STOP Stop button
OUT       M01004	// M_정지 Stop

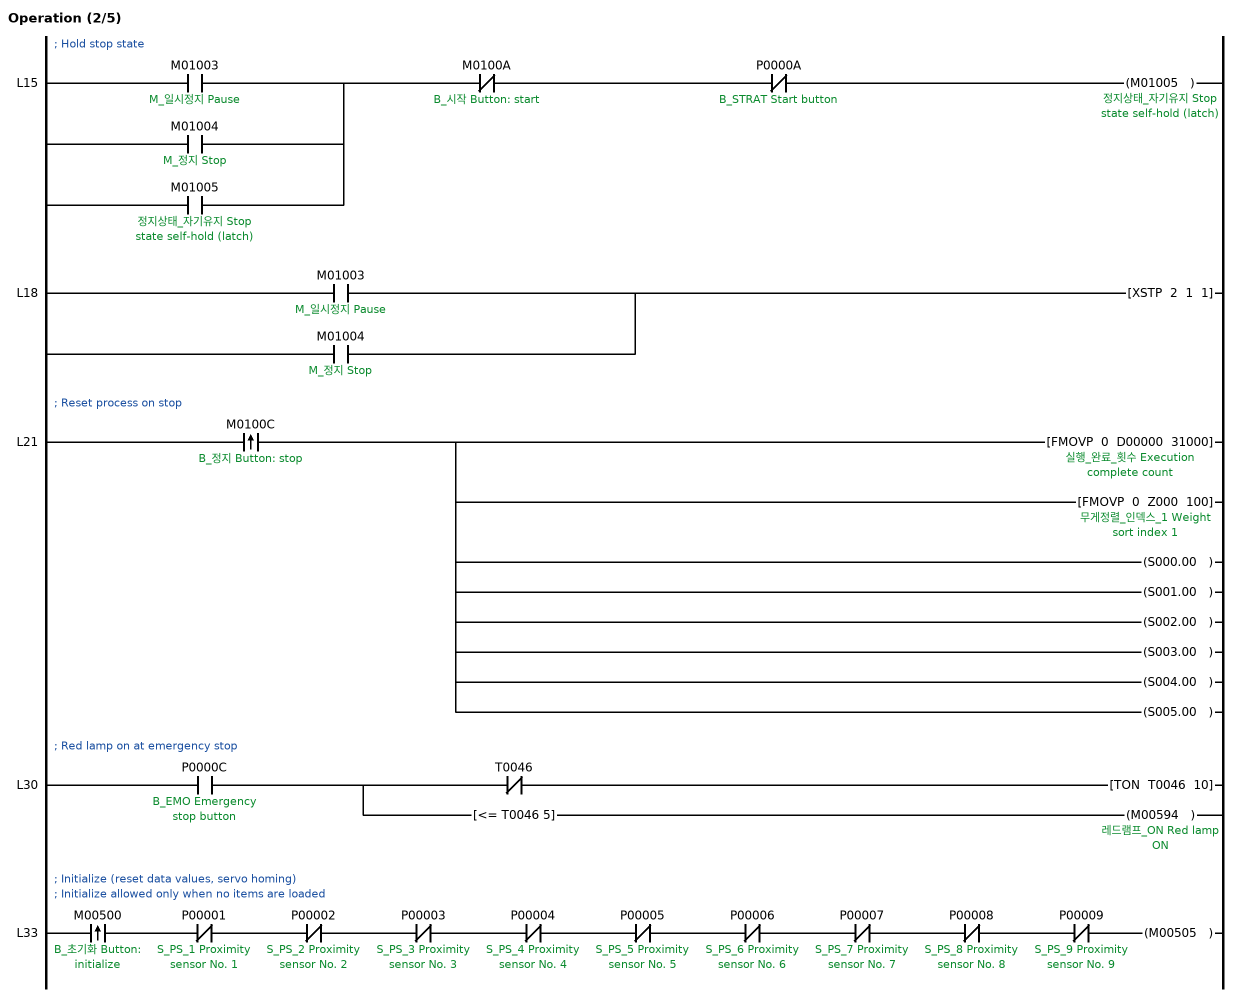
; L15
LOAD      M01003	// M_일시정지 Pause
OR        M01004	// M_정지 Stop
OR        M01005	// 정지상태_자기유지 Stop state self-hold (latch)
AND NOT   M0100A	// B_시작 Button: start
AND NOT   P0000A	// B_STRAT Start button
OUT       M01005	// 정지상태_자기유지 Stop state self-hold (latch)
// output comment: Hold stop state
; L18
LOAD      M01003	// M_일시정지 Pause
OR        M01004	// M_정지 Stop
XSTP      2 1 1
// Reset process on stop
; L21
LOADP     M0100C	// B_정지 Button: stop
FMOVP     0 D00000 31000	// 실행_완료_횟수 Execution complete count
FMOVP     0 Z000 100	// 무게정렬_인덱스_1 Weight sort index 1
OUT       S000.00
OUT       S001.00
OUT       S002.00
OUT       S003.00
OUT       S004.00
OUT       S005.00
// Red lamp on at emergency stop
; L30
LOAD      P0000C	// B_EMO Emergency stop button
MPUSH
AND NOT   T0046
TON       T0046 10
MPOP
AND<=     T0046 5
OUT       M00594	// 레드램프_ON Red lamp ON
// Initialize (reset data values, servo homing)
; L33
LOADP     M00500	// B_초기화 Button: initialize
AND NOT   P00001	// S_PS_1 Proximity sensor No. 1
AND NOT   P00002	// S_PS_2 Proximity sensor No. 2
AND NOT   P00003	// S_PS_3 Proximity sensor No. 3
AND NOT   P00004	// S_PS_4 Proximity sensor No. 4
AND NOT   P00005	// S_PS_5 Proximity sensor No. 5
AND NOT   P00006	// S_PS_6 Proximity sensor No. 6
AND NOT   P00007	// S_PS_7 Proximity sensor No. 7
AND NOT   P00008	// S_PS_8 Proximity sensor No. 8
AND NOT   P00009	// S_PS_9 Proximity sensor No. 9
OUT       M00505
// output comment: Initialize allowed only when no items are loaded

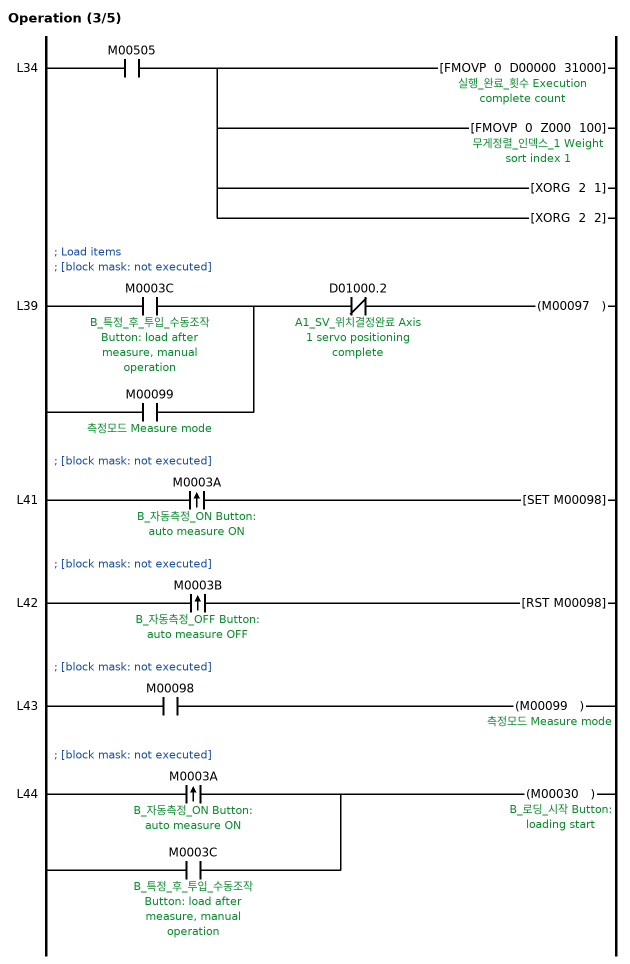
; L34
LOAD      M00505
FMOVP     0 D00000 31000	// 실행_완료_횟수 Execution complete count
FMOVP     0 Z000 100	// 무게정렬_인덱스_1 Weight sort index 1
XORG      2 1
XORG      2 2
// Load items
; L39 (block mask: not executed)
LOAD      M0003C	// B_특정_후_투입_수동조작 Button: load after measure, manual operation
OR        M00099	// 측정모드 Measure mode
AND NOT   D01000.2	// A1_SV_위치결정완료 Axis 1 servo positioning complete
OUT       M00097
; L41 (block mask: not executed)
LOADP     M0003A	// B_자동측정_ON Button: auto measure ON
SET       M00098
; L42 (block mask: not executed)
LOADP     M0003B	// B_자동측정_OFF Button: auto measure OFF
RST       M00098
; L43 (block mask: not executed)
LOAD      M00098
OUT       M00099	// 측정모드 Measure mode
; L44 (block mask: not executed)
LOADP     M0003A	// B_자동측정_ON Button: auto measure ON
OR        M0003C	// B_특정_후_투입_수동조작 Button: load after measure, manual operation
OUT       M00030	// B_로딩_시작 Button: loading start

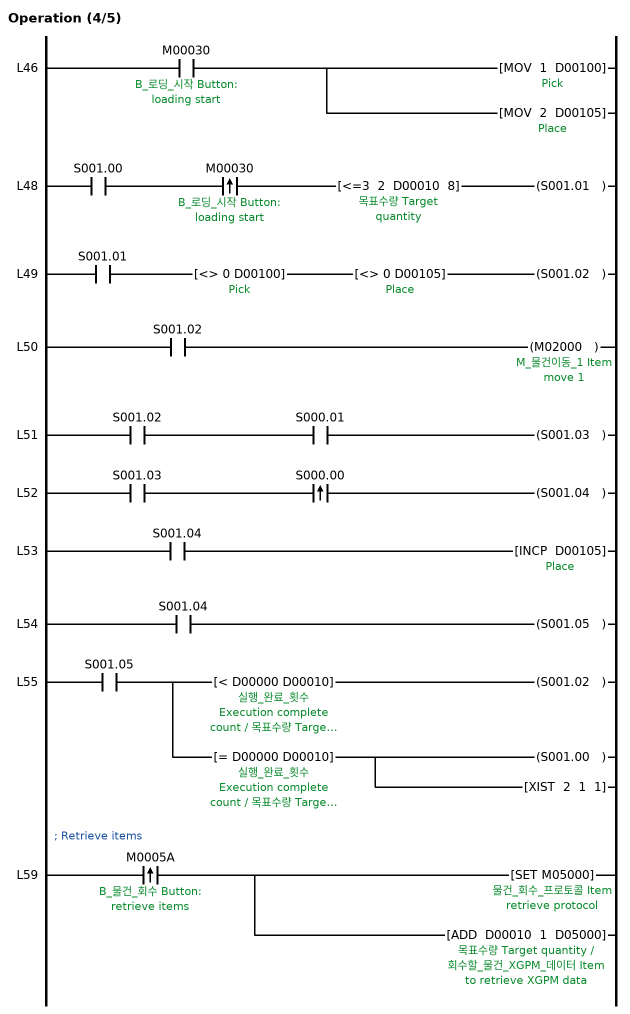
; L46
LOAD      M00030	// B_로딩_시작 Button: loading start
MOV       1 D00100	// Pick
MOV       2 D00105	// Place
; L48
LOAD      S001.00
ANDP      M00030	// B_로딩_시작 Button: loading start
AND<=3    2 D00010 8	// 목표수량 Target quantity
OUT       S001.01
; L49
LOAD      S001.01
AND<>     0 D00100	// Pick
AND<>     0 D00105	// Place
OUT       S001.02
; L50
LOAD      S001.02
OUT       M02000	// M_물건이동_1 Item move 1
; L51
LOAD      S001.02
AND       S000.01
OUT       S001.03
; L52
LOAD      S001.03
ANDP      S000.00
OUT       S001.04
; L53
LOAD      S001.04
INCP      D00105	// Place
; L54
LOAD      S001.04
OUT       S001.05
; L55
LOAD      S001.05
MPUSH
AND<      D00000 D00010	// 실행_완료_횟수 Execution complete count / 목표수량 Target quantity
OUT       S001.02
MPOP
AND=      D00000 D00010	// 실행_완료_횟수 Execution complete count / 목표수량 Target quantity
OUT       S001.00
XIST      2 1 1
// Retrieve items
; L59
LOADP     M0005A	// B_물건_회수 Button: retrieve items
SET       M05000	// 물건_회수_프로토콜 Item retrieve protocol
ADD       D00010 1 D05000	// 목표수량 Target quantity / 회수할_물건_XGPM_데이터 Item to retrieve XGPM data

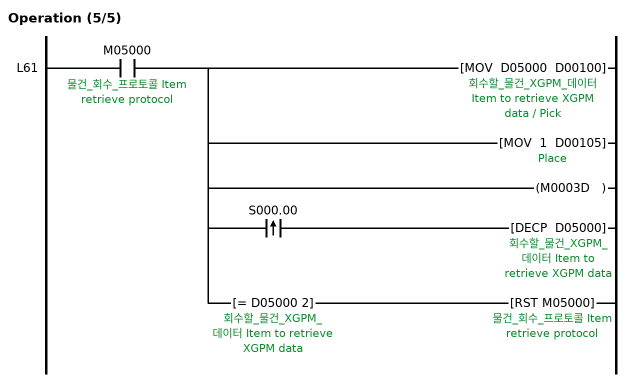
; L61
LOAD      M05000	// 물건_회수_프로토콜 Item retrieve protocol
MOV       D05000 D00100	// 회수할_물건_XGPM_데이터 Item to retrieve XGPM data / Pick
MOV       1 D00105	// Place
OUT       M0003D
MPUSH
ANDP      S000.00
DECP      D05000	// 회수할_물건_XGPM_데이터 Item to retrieve XGPM data
MPOP
AND=      D05000 2	// 회수할_물건_XGPM_데이터 Item to retrieve XGPM data
RST       M05000	// 물건_회수_프로토콜 Item retrieve protocol

PROGRAM Total (task: 스캔 프로그램)

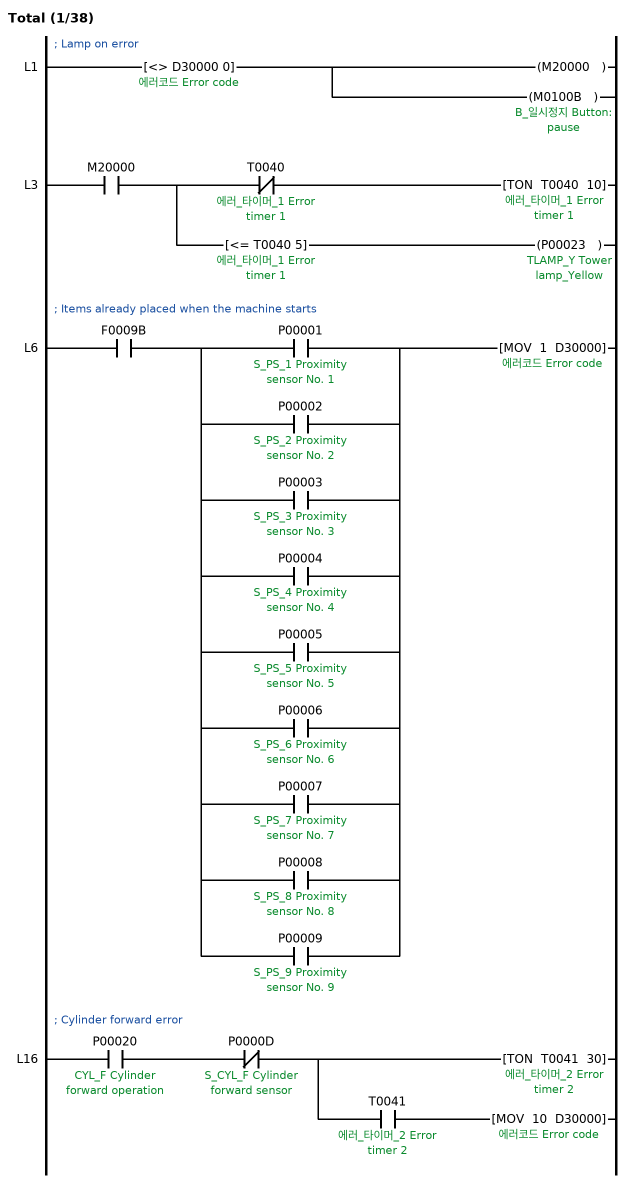
// Lamp on error
; L1
LOAD<>    D30000 0	// 에러코드 Error code
OUT       M20000
OUT       M0100B	// B_일시정지 Button: pause
; L3
LOAD      M20000
MPUSH
AND NOT   T0040	// 에러_타이머_1 Error timer 1
TON       T0040 10	// 에러_타이머_1 Error timer 1
MPOP
AND<=     T0040 5	// 에러_타이머_1 Error timer 1
OUT       P00023	// TLAMP_Y Tower lamp_Yellow
// Items already placed when the machine starts
; L6
LOAD      F0009B
LOAD      P00001	// S_PS_1 Proximity sensor No. 1
OR        P00002	// S_PS_2 Proximity sensor No. 2
OR        P00003	// S_PS_3 Proximity sensor No. 3
OR        P00004	// S_PS_4 Proximity sensor No. 4
OR        P00005	// S_PS_5 Proximity sensor No. 5
OR        P00006	// S_PS_6 Proximity sensor No. 6
OR        P00007	// S_PS_7 Proximity sensor No. 7
OR        P00008	// S_PS_8 Proximity sensor No. 8
OR        P00009	// S_PS_9 Proximity sensor No. 9
AND LOAD
MOV       1 D30000	// 에러코드 Error code
// Cylinder forward error
; L16
LOAD      P00020	// CYL_F Cylinder forward operation
AND NOT   P0000D	// S_CYL_F Cylinder forward sensor
TON       T0041 30	// 에러_타이머_2 Error timer 2
AND       T0041	// 에러_타이머_2 Error timer 2
MOV       10 D30000	// 에러코드 Error code

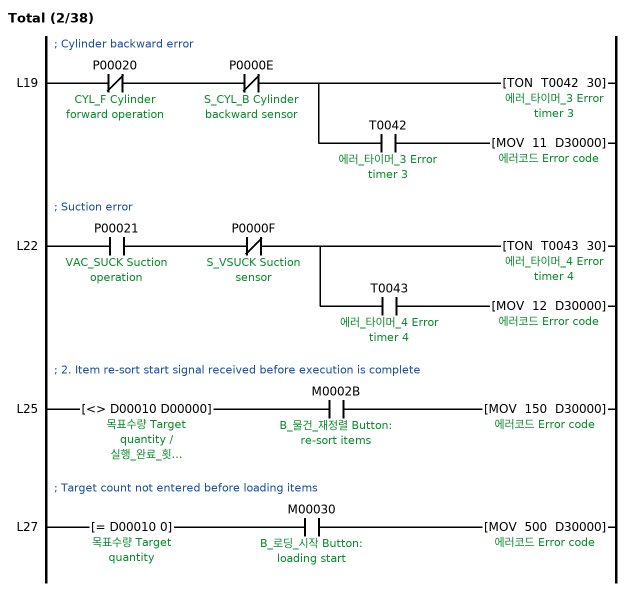
// Cylinder backward error
; L19
LOAD NOT  P00020	// CYL_F Cylinder forward operation
AND NOT   P0000E	// S_CYL_B Cylinder backward sensor
TON       T0042 30	// 에러_타이머_3 Error timer 3
AND       T0042	// 에러_타이머_3 Error timer 3
MOV       11 D30000	// 에러코드 Error code
// Suction error
; L22
LOAD      P00021	// VAC_SUCK Suction operation
AND NOT   P0000F	// S_VSUCK Suction sensor
TON       T0043 30	// 에러_타이머_4 Error timer 4
AND       T0043	// 에러_타이머_4 Error timer 4
MOV       12 D30000	// 에러코드 Error code
// 2. Item re-sort start signal received before execution is complete
; L25
LOAD<>    D00010 D00000	// 목표수량 Target quantity / 실행_완료_횟수 Execution complete count
AND       M0002B	// B_물건_재정렬 Button: re-sort items
MOV       150 D30000	// 에러코드 Error code
// Target count not entered before loading items
; L27
LOAD=     D00010 0	// 목표수량 Target quantity
AND       M00030	// B_로딩_시작 Button: loading start
MOV       500 D30000	// 에러코드 Error code

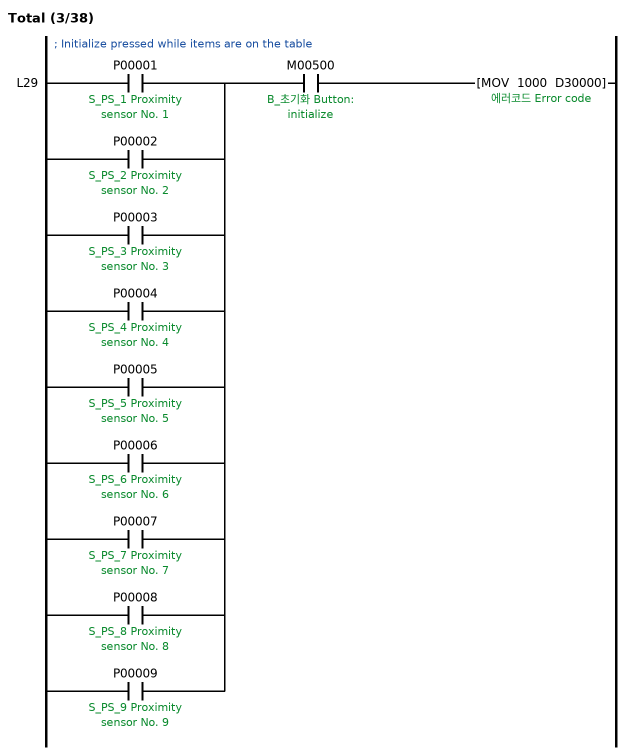
// Initialize pressed while items are on the table
; L29
LOAD      P00001	// S_PS_1 Proximity sensor No. 1
OR        P00002	// S_PS_2 Proximity sensor No. 2
OR        P00003	// S_PS_3 Proximity sensor No. 3
OR        P00004	// S_PS_4 Proximity sensor No. 4
OR        P00005	// S_PS_5 Proximity sensor No. 5
OR        P00006	// S_PS_6 Proximity sensor No. 6
OR        P00007	// S_PS_7 Proximity sensor No. 7
OR        P00008	// S_PS_8 Proximity sensor No. 8
OR        P00009	// S_PS_9 Proximity sensor No. 9
AND       M00500	// B_초기화 Button: initialize
MOV       1000 D30000	// 에러코드 Error code

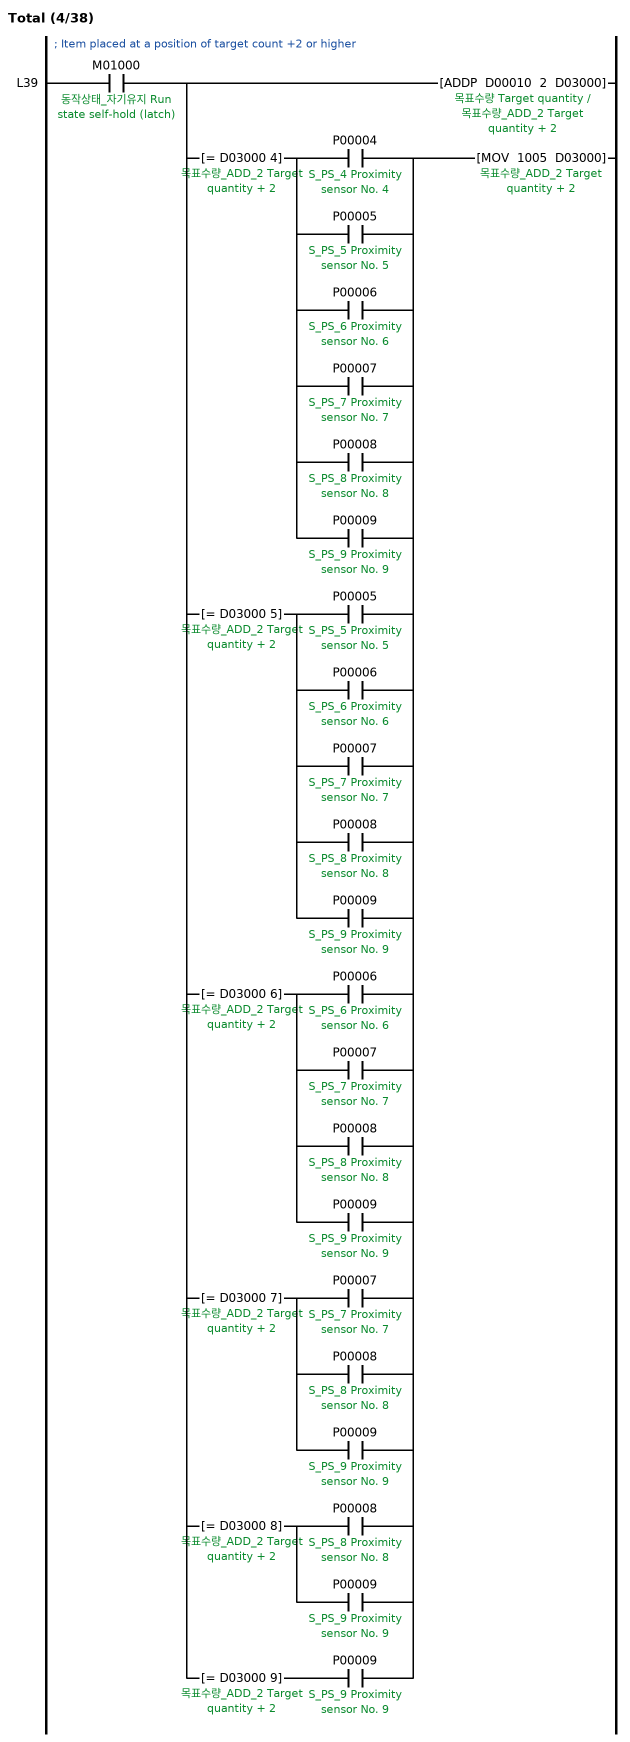
// Item placed at a position of target count +2 or higher
; L39
LOAD      M01000	// 동작상태_자기유지 Run state self-hold (latch)
ADDP      D00010 2 D03000	// 목표수량 Target quantity / 목표수량_ADD_2 Target quantity + 2
LOAD=     D03000 4	// 목표수량_ADD_2 Target quantity + 2
LOAD      P00004	// S_PS_4 Proximity sensor No. 4
OR        P00005	// S_PS_5 Proximity sensor No. 5
OR        P00006	// S_PS_6 Proximity sensor No. 6
OR        P00007	// S_PS_7 Proximity sensor No. 7
OR        P00008	// S_PS_8 Proximity sensor No. 8
OR        P00009	// S_PS_9 Proximity sensor No. 9
AND LOAD
LOAD=     D03000 5	// 목표수량_ADD_2 Target quantity + 2
LOAD      P00005	// S_PS_5 Proximity sensor No. 5
OR        P00006	// S_PS_6 Proximity sensor No. 6
OR        P00007	// S_PS_7 Proximity sensor No. 7
OR        P00008	// S_PS_8 Proximity sensor No. 8
OR        P00009	// S_PS_9 Proximity sensor No. 9
AND LOAD
OR LOAD
LOAD=     D03000 6	// 목표수량_ADD_2 Target quantity + 2
LOAD      P00006	// S_PS_6 Proximity sensor No. 6
OR        P00007	// S_PS_7 Proximity sensor No. 7
OR        P00008	// S_PS_8 Proximity sensor No. 8
OR        P00009	// S_PS_9 Proximity sensor No. 9
AND LOAD
OR LOAD
LOAD=     D03000 7	// 목표수량_ADD_2 Target quantity + 2
LOAD      P00007	// S_PS_7 Proximity sensor No. 7
OR        P00008	// S_PS_8 Proximity sensor No. 8
OR        P00009	// S_PS_9 Proximity sensor No. 9
AND LOAD
OR LOAD
LOAD=     D03000 8	// 목표수량_ADD_2 Target quantity + 2
LOAD      P00008	// S_PS_8 Proximity sensor No. 8
OR        P00009	// S_PS_9 Proximity sensor No. 9
AND LOAD
OR LOAD
LOAD=     D03000 9	// 목표수량_ADD_2 Target quantity + 2
AND       P00009	// S_PS_9 Proximity sensor No. 9
OR LOAD
AND LOAD
MOV       1005 D03000	// 목표수량_ADD_2 Target quantity + 2

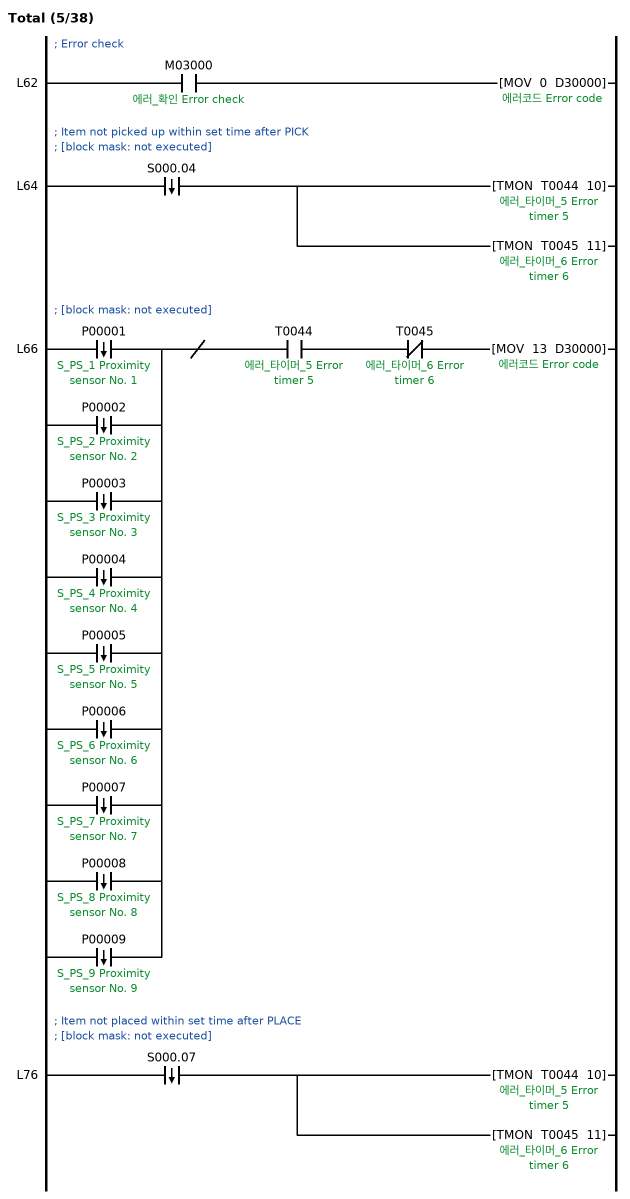
// Error check
; L62
LOAD      M03000	// 에러_확인 Error check
MOV       0 D30000	// 에러코드 Error code
// Item not picked up within set time after PICK
; L64 (block mask: not executed)
LOADN     S000.04
TMON      T0044 10	// 에러_타이머_5 Error timer 5
TMON      T0045 11	// 에러_타이머_6 Error timer 6
; L66 (block mask: not executed)
LOADN     P00001	// S_PS_1 Proximity sensor No. 1
ORN       P00002	// S_PS_2 Proximity sensor No. 2
ORN       P00003	// S_PS_3 Proximity sensor No. 3
ORN       P00004	// S_PS_4 Proximity sensor No. 4
ORN       P00005	// S_PS_5 Proximity sensor No. 5
ORN       P00006	// S_PS_6 Proximity sensor No. 6
ORN       P00007	// S_PS_7 Proximity sensor No. 7
ORN       P00008	// S_PS_8 Proximity sensor No. 8
ORN       P00009	// S_PS_9 Proximity sensor No. 9
NOT
AND       T0044	// 에러_타이머_5 Error timer 5
AND NOT   T0045	// 에러_타이머_6 Error timer 6
MOV       13 D30000	// 에러코드 Error code
// Item not placed within set time after PLACE
; L76 (block mask: not executed)
LOADN     S000.07
TMON      T0044 10	// 에러_타이머_5 Error timer 5
TMON      T0045 11	// 에러_타이머_6 Error timer 6

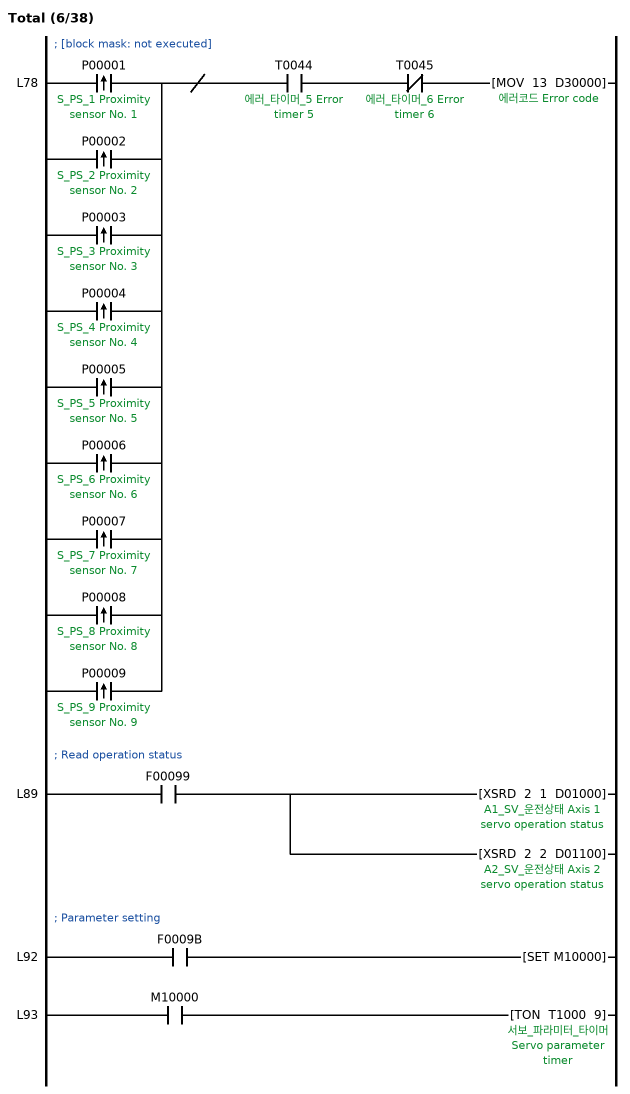
; L78 (block mask: not executed)
LOADP     P00001	// S_PS_1 Proximity sensor No. 1
ORP       P00002	// S_PS_2 Proximity sensor No. 2
ORP       P00003	// S_PS_3 Proximity sensor No. 3
ORP       P00004	// S_PS_4 Proximity sensor No. 4
ORP       P00005	// S_PS_5 Proximity sensor No. 5
ORP       P00006	// S_PS_6 Proximity sensor No. 6
ORP       P00007	// S_PS_7 Proximity sensor No. 7
ORP       P00008	// S_PS_8 Proximity sensor No. 8
ORP       P00009	// S_PS_9 Proximity sensor No. 9
NOT
AND       T0044	// 에러_타이머_5 Error timer 5
AND NOT   T0045	// 에러_타이머_6 Error timer 6
MOV       13 D30000	// 에러코드 Error code
// Read operation status
; L89
LOAD      F00099
XSRD      2 1 D01000	// A1_SV_운전상태 Axis 1 servo operation status
XSRD      2 2 D01100	// A2_SV_운전상태 Axis 2 servo operation status
// Parameter setting
; L92
LOAD      F0009B
SET       M10000
; L93
LOAD      M10000
TON       T1000 9	// 서보_파라미터_타이머 Servo parameter timer

